</description>
*)
{endregion}
FUNCTION_BLOCK AssertInTimespan_LDT EXTENDS AssertionBase
VAR_INPUT
    IN : LDT; //! Actual value checked or observed by this Assertion.
    StartTime : LDT; //! Inclusive start of the time span; must not exceed EndTime.
    EndTime : LDT; //! Inclusive end of the time span; must not precede StartTime.
END_VAR

SUPER^();

{region 'Documentation'}
(*!
<summary>Evaluate the typed temporal relation and report higher-priority errors first.</summary>
*)
{endregion}
METHOD PROTECTED Assert
VAR
    Message : STRING(GVL_Constants.MessageLength);
    StartTimeText : STRING(GVL_Constants.AssertionValueLength);
    EndTimeText : STRING(GVL_Constants.AssertionValueLength);
    ActualText : STRING(GVL_Constants.AssertionValueLength);
END_VAR
IF NOT EvaluationActive THEN
    RETURN;
END_IF;

IF Result = E_Result.Error THEN
    RETURN;
END_IF;

IF StartTime > EndTime THEN
    StartTimeText := LDT_TO_STRING(StartTime);
    EndTimeText := LDT_TO_STRING(EndTime);
    Message := CONCAT('Assertion error: start time exceeds end time. StartTime = ',
        StartTimeText);
    Message := CONCAT(Message, ', EndTime = ');
    Message := CONCAT(Message, EndTimeText);
    Message := CONCAT(Message, '.');
    Error(Message := Message);
    RETURN;
END_IF;

IF Result = E_Result.Failed THEN
    RETURN;
END_IF;

IF (IN < StartTime) OR (IN > EndTime) THEN
    StartTimeText := LDT_TO_STRING(StartTime);
    EndTimeText := LDT_TO_STRING(EndTime);
    ActualText := LDT_TO_STRING(IN);
    Message := CONCAT('Assertion failed: value is outside allowed timespan. StartTime = ',
        StartTimeText);
    Message := CONCAT(Message, ', EndTime = ');
    Message := CONCAT(Message, EndTimeText);
    Message := CONCAT(Message, ', Actual = ');
    Message := CONCAT(Message, ActualText);
    Message := CONCAT(Message, '.');
    Fail(Message := Message);
    RETURN;
END_IF;

Pass();
END_METHOD

END_FUNCTION_BLOCK

// ---- Framework/Assertions/POU/BasicTypes/LDT/AssertLaterThan_LDT.TcPOU
{region 'Documentation'}
(*!
<summary>Check that IN is strictly later than Minimum.</summary>
*)
{endregion}
FUNCTION_BLOCK AssertLaterThan_LDT EXTENDS AssertionBase
VAR_INPUT
    IN : LDT; //! Actual value checked or observed by this Assertion.
    Minimum : LDT; //! Exclusive lower bound; the actual value or count must be greater.
END_VAR

SUPER^();

{region 'Documentation'}
(*!
<summary>Evaluate the typed temporal relation and report higher-priority errors first.</summary>
*)
{endregion}
METHOD PROTECTED Assert
VAR
    Message : STRING(GVL_Constants.MessageLength);
    MinimumText : STRING(GVL_Constants.AssertionValueLength);
    ActualText : STRING(GVL_Constants.AssertionValueLength);
END_VAR
IF NOT EvaluationActive THEN
    RETURN;
END_IF;

IF Result = E_Result.Error THEN
    RETURN;
END_IF;

IF Result = E_Result.Failed THEN
    RETURN;
END_IF;

IF IN <= Minimum THEN
    MinimumText := LDT_TO_STRING(Minimum);
    ActualText := LDT_TO_STRING(IN);
    Message := CONCAT('Assertion failed: value is not later than limit. Minimum = ',
        MinimumText);
    Message := CONCAT(Message, ', Actual = ');
    Message := CONCAT(Message, ActualText);
    Message := CONCAT(Message, '.');
    Fail(Message := Message);
    RETURN;
END_IF;

Pass();
END_METHOD

END_FUNCTION_BLOCK

// ---- Framework/Assertions/POU/BasicTypes/LDT/AssertNotEqual_LDT.TcPOU
{region 'Documentation'}
(*!
<summary>Checks inequality with the forbidden LDT value.</summary>
*)
{endregion}
FUNCTION_BLOCK AssertNotEqual_LDT EXTENDS AssertionBase
VAR_INPUT
    IN : LDT; //! Actual value checked or observed by this Assertion.
    Expected : LDT; //! Value that must differ from IN under this Assertion's comparison rules.
END_VAR

SUPER^();

{region 'Documentation'}
(*!
<summary>Evaluate the typed temporal relation and report higher-priority errors first.</summary>
*)
{endregion}
METHOD PROTECTED Assert
VAR
    Message : STRING(GVL_Constants.MessageLength);
    ExpectedText : STRING(GVL_Constants.AssertionValueLength);
    ActualText : STRING(GVL_Constants.AssertionValueLength);
END_VAR
IF NOT EvaluationActive THEN
    RETURN;
END_IF;

IF Result = E_Result.Error THEN
    RETURN;
END_IF;

IF Result = E_Result.Failed THEN
    RETURN;
END_IF;

IF IN = Expected THEN
    ExpectedText := LDT_TO_STRING(Expected);
    ActualText := LDT_TO_STRING(IN);
    Message := CONCAT('Assertion failed: values are equal but should differ. NotExpected = ',
        ExpectedText);
    Message := CONCAT(Message, ', Actual = ');
    Message := CONCAT(Message, ActualText);
    Message := CONCAT(Message, '.');
    Fail(Message := Message);
    RETURN;
END_IF;

Pass();
END_METHOD

END_FUNCTION_BLOCK

// ---- Framework/Assertions/POU/BasicTypes/LDT/AssertNotInTimespan_LDT.TcPOU
{region 'Documentation'}
(*!
<summary>Check that IN is outside the inclusive StartTime..EndTime interval.</summary>
<description>

StartTime &gt; EndTime reports Error during active evaluation; equal bounds are
valid.

</description>
*)
{endregion}
FUNCTION_BLOCK AssertNotInTimespan_LDT EXTENDS AssertionBase
VAR_INPUT
    IN : LDT; //! Actual value checked or observed by this Assertion.
    StartTime : LDT; //! Inclusive start of the time span; must not exceed EndTime.
    EndTime : LDT; //! Inclusive end of the time span; must not precede StartTime.
END_VAR

SUPER^();

{region 'Documentation'}
(*!
<summary>Evaluate the typed temporal relation and report higher-priority errors first.</summary>
*)
{endregion}
METHOD PROTECTED Assert
VAR
    Message : STRING(GVL_Constants.MessageLength);
    StartTimeText : STRING(GVL_Constants.AssertionValueLength);
    EndTimeText : STRING(GVL_Constants.AssertionValueLength);
    ActualText : STRING(GVL_Constants.AssertionValueLength);
END_VAR
IF NOT EvaluationActive THEN
    RETURN;
END_IF;

IF Result = E_Result.Error THEN
    RETURN;
END_IF;

IF StartTime > EndTime THEN
    StartTimeText := LDT_TO_STRING(StartTime);
    EndTimeText := LDT_TO_STRING(EndTime);
    Message := CONCAT('Assertion error: start time exceeds end time. StartTime = ',
        StartTimeText);
    Message := CONCAT(Message, ', EndTime = ');
    Message := CONCAT(Message, EndTimeText);
    Message := CONCAT(Message, '.');
    Error(Message := Message);
    RETURN;
END_IF;

IF Result = E_Result.Failed THEN
    RETURN;
END_IF;

IF (IN >= StartTime) AND (IN <= EndTime) THEN
    StartTimeText := LDT_TO_STRING(StartTime);
    EndTimeText := LDT_TO_STRING(EndTime);
    ActualText := LDT_TO_STRING(IN);
    Message := CONCAT('Assertion failed: value is inside forbidden timespan. StartTime = ',
        StartTimeText);
    Message := CONCAT(Message, ', EndTime = ');
    Message := CONCAT(Message, EndTimeText);
    Message := CONCAT(Message, ', Actual = ');
    Message := CONCAT(Message, ActualText);
    Message := CONCAT(Message, '.');
    Fail(Message := Message);
    RETURN;
END_IF;

Pass();
END_METHOD

END_FUNCTION_BLOCK

// ---- Framework/Assertions/POU/BasicTypes/LDT/AssertNoValueChange_LDT.TcPOU
{region 'Documentation'}
(*!
<summary>Check equality between consecutive active observations.</summary>
<description>

The first active observation establishes a baseline without deciding a result. Disabling
observation invalidates that baseline, not the held Result. Re-enabling first establishes a new
baseline; Reset clears history.

ObserveFirstCycle FALSE delays the first observation by one enabled call.

</description>
*)
{endregion}
FUNCTION_BLOCK AssertNoValueChange_LDT EXTENDS AssertionBase
VAR_INPUT
    IN : LDT; //! Actual value to observe.
END_VAR
VAR
    FINPrevious : LDT;
    FObservationPrevious : BOOL;
    FEvaluationActive : BOOL;
END_VAR

SUPER^();

{region 'Documentation'}
(*!
<summary>Observe the current value before evaluating a change against the previous observation.</summary>
*)
{endregion}
METHOD PROTECTED Assert
VAR
    PreviousValue : LDT;
    Message : STRING(GVL_Constants.MessageLength);
    PreviousText : STRING(GVL_Constants.AssertionValueLength);
    ActualText : STRING(GVL_Constants.AssertionValueLength);
END_VAR
FEvaluationActive := ObservationActive AND FObservationPrevious;
FObservationPrevious := ObservationActive;

IF NOT ObservationActive THEN
    RETURN;
END_IF;

PreviousValue := FINPrevious;
FINPrevious := IN;

IF NOT EvaluationActive THEN
    RETURN;
END_IF;

IF Result = E_Result.Error THEN
    RETURN;
END_IF;

IF Result = E_Result.Failed THEN
    RETURN;
END_IF;

IF IN <> PreviousValue THEN
    PreviousText := LDT_TO_STRING(PreviousValue);
    ActualText := LDT_TO_STRING(IN);
    Message := CONCAT('Assertion failed: value changed unexpectedly. Previous = ',
        PreviousText);
    Message := CONCAT(Message, ', Actual = ');
    Message := CONCAT(Message, ActualText);
    Message := CONCAT(Message, '.');
    Fail(Message := Message);
    RETURN;
END_IF;

Pass();
END_METHOD

{region 'Documentation'}
(*!
<summary>Current/last call has an active observation and a preceding observation
baseline.</summary>
*)
{endregion}
{attribute 'monitoring' := 'call'}
PROPERTY PUBLIC EvaluationActive : BOOL //! Current/last call has an active observation and a preceding observation baseline.
GET // PUBLIC
EvaluationActive := FEvaluationActive;
END_GET
END_PROPERTY

{region 'Documentation'}
(*!
<summary>Clear observation history and the current evaluation gate.</summary>
*)
{endregion}
METHOD PROTECTED ResetAssertion
FINPrevious := LDT#1970-01-01-00:00:00;
FObservationPrevious := FALSE;
FEvaluationActive := FALSE;
END_METHOD

END_FUNCTION_BLOCK

// ---- Framework/Assertions/POU/BasicTypes/LInt/AssertNoValueChange_LInt.TcPOU
{region 'Documentation'}
(*!
<summary>Check equality between consecutive active observations.</summary>
<description>

The first active observation establishes a baseline without deciding a result. Disabling
observation invalidates that baseline, not the held Result. Re-enabling first establishes a new
baseline; Reset clears history.

ObserveFirstCycle FALSE delays the first observation by one enabled call.

</description>
*)
{endregion}
FUNCTION_BLOCK AssertNoValueChange_LInt EXTENDS AssertionBase
VAR_INPUT
    IN : LINT; //! Actual value to observe.
END_VAR
VAR
    FINPrevious : LINT;
    FObservationPrevious : BOOL;
    FEvaluationActive : BOOL;
END_VAR

SUPER^();

{region 'Documentation'}
(*!
<summary>Observe the current value before evaluating a change against the previous observation.</summary>
*)
{endregion}
METHOD PROTECTED Assert
VAR
    PreviousValue : LINT;
    Message : STRING(GVL_Constants.MessageLength);
    PreviousText : STRING(GVL_Constants.AssertionValueLength);
    ActualText : STRING(GVL_Constants.AssertionValueLength);
END_VAR
FEvaluationActive := ObservationActive AND FObservationPrevious;
FObservationPrevious := ObservationActive;

IF NOT ObservationActive THEN
    RETURN;
END_IF;

PreviousValue := FINPrevious;
FINPrevious := IN;

IF NOT EvaluationActive THEN
    RETURN;
END_IF;

IF Result = E_Result.Error THEN
    RETURN;
END_IF;

IF Result = E_Result.Failed THEN
    RETURN;
END_IF;

IF IN <> PreviousValue THEN
    PreviousText := LINT_TO_STRING(PreviousValue);
    ActualText := LINT_TO_STRING(IN);
    Message := CONCAT('Assertion failed: value changed unexpectedly. Previous = ',
        PreviousText);
    Message := CONCAT(Message, ', Actual = ');
    Message := CONCAT(Message, ActualText);
    Message := CONCAT(Message, '.');
    Fail(Message := Message);
    RETURN;
END_IF;

Pass();
END_METHOD

{region 'Documentation'}
(*!
<summary>Current/last call has an active observation and a preceding observation
baseline.</summary>
*)
{endregion}
{attribute 'monitoring' := 'call'}
PROPERTY PUBLIC EvaluationActive : BOOL //! Current/last call has an active observation and a preceding observation baseline.
GET // PUBLIC
EvaluationActive := FEvaluationActive;
END_GET
END_PROPERTY

{region 'Documentation'}
(*!
<summary>Clear observation history and the current evaluation gate.</summary>
*)
{endregion}
METHOD PROTECTED ResetAssertion
FINPrevious := 0;
FObservationPrevious := FALSE;
FEvaluationActive := FALSE;
END_METHOD

END_FUNCTION_BLOCK

// ---- Framework/Assertions/POU/BasicTypes/LInt/AssertSequence_LInt.TcPOU
{region 'Documentation'}
(*!
<summary>Checks the observed value sequence; Evaluate also checks the current value and
completeness.</summary>
<description>

Uses the whole Expected array from its declared lower bound. Keep its binding, bounds and
values stable until Reset; supply it on reset and disabled FB calls as well.

Observation accepts the current expected value and then permits advancing by one element
on a later change. Repeated equal values do not advance. An unexpected value or an out-of-range
sequence index reports Failed.

Evaluate checks the current value and requires the final expected element to have been
reached; only then can the result become Passed. Disabling observation retains progression.
Reset restarts it.

</description>
*)
{endregion}
FUNCTION_BLOCK AssertSequence_LInt EXTENDS AssertionWithEvaluationBase
VAR_INPUT
    IN : LINT; //! Actual value to observe.
END_VAR
VAR_IN_OUT CONSTANT
    Expected : ARRAY[*] OF LINT; //! Complete expected sequence; read without modifying the supplied array.
END_VAR
VAR
    FExpectedIndex : DINT;
    FSequenceIndexInitialized : BOOL;
    FAllowAdvance : BOOL;
END_VAR

SUPER^();

{region 'Documentation'}
(*!
<summary>Advances at most one entry and checks the current value before explicit completeness evaluation.</summary>
*)
{endregion}
METHOD PROTECTED Assert
VAR
    LowerIndex : DINT;
    UpperIndex : DINT;
    ExpectedValue : LINT;
    MatchesExpected : BOOL;
    AllowAdvance : BOOL;
    Message : STRING(GVL_Constants.MessageLength);
    ExpectedText : STRING(GVL_Constants.AssertionValueLength);
    ActualText : STRING(GVL_Constants.AssertionValueLength);
END_VAR
LowerIndex := LOWER_BOUND(Expected, 1);
UpperIndex := UPPER_BOUND(Expected, 1);

IF NOT FSequenceIndexInitialized THEN
    FExpectedIndex := LowerIndex;
    FSequenceIndexInitialized := TRUE;
END_IF;

IF NOT (ObservationActive OR EvaluationActive) THEN
    RETURN;
END_IF;

IF Result = E_Result.Error THEN
    RETURN;
END_IF;

IF Result = E_Result.Failed THEN
    RETURN;
END_IF;

IF (FExpectedIndex < LowerIndex) OR (FExpectedIndex > UpperIndex) THEN
    Message := CONCAT('Assertion failed: sequence index out of range. ExpectedIndex = ',
        DINT_TO_STRING(FExpectedIndex));
    Message := CONCAT(Message, ', LowerIndex = ');
    Message := CONCAT(Message, DINT_TO_STRING(LowerIndex));
    Message := CONCAT(Message, ', UpperIndex = ');
    Message := CONCAT(Message, DINT_TO_STRING(UpperIndex));
    Message := CONCAT(Message, '.');
    Fail(Message := Message);
    RETURN;
END_IF;

AllowAdvance := FAllowAdvance;
IF ObservationActive THEN
    FAllowAdvance := TRUE;
END_IF;

ExpectedValue := Expected[FExpectedIndex];
MatchesExpected := IN = ExpectedValue;

IF AllowAdvance AND NOT MatchesExpected THEN
    IF FExpectedIndex = UpperIndex THEN
        Message := CONCAT('Assertion failed: sequence continued beyond its last entry. LastIndex = ',
            DINT_TO_STRING(UpperIndex));
        Message := CONCAT(Message, '.');
        Fail(Message := Message);
        RETURN;
    END_IF;

    FExpectedIndex := FExpectedIndex + 1;
    ExpectedValue := Expected[FExpectedIndex];
    MatchesExpected := IN = ExpectedValue;
END_IF;

IF NOT MatchesExpected THEN
    ExpectedText := LINT_TO_STRING(ExpectedValue);
    ActualText := LINT_TO_STRING(IN);
    Message := CONCAT('Assertion failed: sequence value does not match. ExpectedIndex = ',
        DINT_TO_STRING(FExpectedIndex));
    Message := CONCAT(Message, ', Expected = ');
    Message := CONCAT(Message, ExpectedText);
    Message := CONCAT(Message, ', Actual = ');
    Message := CONCAT(Message, ActualText);
    Message := CONCAT(Message, '.');
    Fail(Message := Message);
    RETURN;
END_IF;

IF NOT EvaluationActive THEN
    RETURN;
END_IF;

IF FExpectedIndex <> UpperIndex THEN
    Message := CONCAT('Assertion failed: sequence is incomplete. ExpectedIndex = ',
        DINT_TO_STRING(FExpectedIndex));
    Message := CONCAT(Message, ', LastIndex = ');
    Message := CONCAT(Message, DINT_TO_STRING(UpperIndex));
    Message := CONCAT(Message, '.');
    Fail(Message := Message);
    RETURN;
END_IF;

Pass();
END_METHOD

{region 'Documentation'}
(*!
<summary>Restart progression at the bound Expected array's lower index.</summary>
<description>

Runs only during the reset FB call with Expected supplied, not directly from Reset or
Initialize. Clears permission to advance from a previous observation.

</description>
*)
{endregion}
METHOD PROTECTED ResetAssertion
FExpectedIndex := LOWER_BOUND(Expected, 1);
FSequenceIndexInitialized := TRUE;
FAllowAdvance := FALSE;
END_METHOD

END_FUNCTION_BLOCK

// ---- Framework/Assertions/POU/BasicTypes/LTime/AssertEarlierThan_LTime.TcPOU
{region 'Documentation'}
(*!
<summary>Check that IN is strictly earlier than Maximum.</summary>
*)
{endregion}
FUNCTION_BLOCK AssertEarlierThan_LTime EXTENDS AssertionBase
VAR_INPUT
    IN : LTIME; //! Actual value checked or observed by this Assertion.
    Maximum : LTIME; //! Exclusive upper bound; the actual value or count must be smaller.
END_VAR

SUPER^();

{region 'Documentation'}
(*!
<summary>Evaluate the typed duration relation and report higher-priority errors first.</summary>
*)
{endregion}
METHOD PROTECTED Assert
VAR
    Message : STRING(GVL_Constants.MessageLength);
    MaximumText : STRING(GVL_Constants.AssertionValueLength);
    ActualText : STRING(GVL_Constants.AssertionValueLength);
END_VAR
IF NOT EvaluationActive THEN
    RETURN;
END_IF;

IF Result = E_Result.Error THEN
    RETURN;
END_IF;

IF Result = E_Result.Failed THEN
    RETURN;
END_IF;

IF IN >= Maximum THEN
    MaximumText := LTIME_TO_STRING(Maximum);
    ActualText := LTIME_TO_STRING(IN);
    Message := CONCAT('Assertion failed: value is not earlier than limit. Maximum = ',
        MaximumText);
    Message := CONCAT(Message, ', Actual = ');
    Message := CONCAT(Message, ActualText);
    Message := CONCAT(Message, '.');
    Fail(Message := Message);
    RETURN;
END_IF;

Pass();
END_METHOD

END_FUNCTION_BLOCK

// ---- Framework/Assertions/POU/BasicTypes/LTime/AssertInTimespan_LTime.TcPOU
{region 'Documentation'}
(*!
<summary>Check that IN is inside the inclusive StartTime..EndTime interval.</summary>
<description>

StartTime &gt; EndTime reports Error during active evaluation; equal bounds are
valid.

</description>
*)
{endregion}
FUNCTION_BLOCK AssertInTimespan_LTime EXTENDS AssertionBase
VAR_INPUT
    IN : LTIME; //! Actual value checked or observed by this Assertion.
    StartTime : LTIME; //! Inclusive start of the time span; must not exceed EndTime.
    EndTime : LTIME; //! Inclusive end of the time span; must not precede StartTime.
END_VAR

SUPER^();

{region 'Documentation'}
(*!
<summary>Evaluate the typed duration relation and report higher-priority errors first.</summary>
*)
{endregion}
METHOD PROTECTED Assert
VAR
    Message : STRING(GVL_Constants.MessageLength);
    StartTimeText : STRING(GVL_Constants.AssertionValueLength);
    EndTimeText : STRING(GVL_Constants.AssertionValueLength);
    ActualText : STRING(GVL_Constants.AssertionValueLength);
END_VAR
IF NOT EvaluationActive THEN
    RETURN;
END_IF;

IF Result = E_Result.Error THEN
    RETURN;
END_IF;

IF StartTime > EndTime THEN
    StartTimeText := LTIME_TO_STRING(StartTime);
    EndTimeText := LTIME_TO_STRING(EndTime);
    Message := CONCAT('Assertion error: start time exceeds end time. StartTime = ',
        StartTimeText);
    Message := CONCAT(Message, ', EndTime = ');
    Message := CONCAT(Message, EndTimeText);
    Message := CONCAT(Message, '.');
    Error(Message := Message);
    RETURN;
END_IF;

IF Result = E_Result.Failed THEN
    RETURN;
END_IF;

IF (IN < StartTime) OR (IN > EndTime) THEN
    StartTimeText := LTIME_TO_STRING(StartTime);
    EndTimeText := LTIME_TO_STRING(EndTime);
    ActualText := LTIME_TO_STRING(IN);
    Message := CONCAT('Assertion failed: value is outside allowed timespan. StartTime = ',
        StartTimeText);
    Message := CONCAT(Message, ', EndTime = ');
    Message := CONCAT(Message, EndTimeText);
    Message := CONCAT(Message, ', Actual = ');
    Message := CONCAT(Message, ActualText);
    Message := CONCAT(Message, '.');
    Fail(Message := Message);
    RETURN;
END_IF;

Pass();
END_METHOD

END_FUNCTION_BLOCK

// ---- Framework/Assertions/POU/BasicTypes/LTime/AssertLaterThan_LTime.TcPOU
{region 'Documentation'}
(*!
<summary>Check that IN is strictly later than Minimum.</summary>
*)
{endregion}
FUNCTION_BLOCK AssertLaterThan_LTime EXTENDS AssertionBase
VAR_INPUT
    IN : LTIME; //! Actual value checked or observed by this Assertion.
    Minimum : LTIME; //! Exclusive lower bound; the actual value or count must be greater.
END_VAR

SUPER^();

{region 'Documentation'}
(*!
<summary>Evaluate the typed duration relation and report higher-priority errors first.</summary>
*)
{endregion}
METHOD PROTECTED Assert
VAR
    Message : STRING(GVL_Constants.MessageLength);
    MinimumText : STRING(GVL_Constants.AssertionValueLength);
    ActualText : STRING(GVL_Constants.AssertionValueLength);
END_VAR
IF NOT EvaluationActive THEN
    RETURN;
END_IF;

IF Result = E_Result.Error THEN
    RETURN;
END_IF;

IF Result = E_Result.Failed THEN
    RETURN;
END_IF;

IF IN <= Minimum THEN
    MinimumText := LTIME_TO_STRING(Minimum);
    ActualText := LTIME_TO_STRING(IN);
    Message := CONCAT('Assertion failed: value is not later than limit. Minimum = ',
        MinimumText);
    Message := CONCAT(Message, ', Actual = ');
    Message := CONCAT(Message, ActualText);
    Message := CONCAT(Message, '.');
    Fail(Message := Message);
    RETURN;
END_IF;

Pass();
END_METHOD

END_FUNCTION_BLOCK

// ---- Framework/Assertions/POU/BasicTypes/LTime/AssertNotEqual_LTime.TcPOU
{region 'Documentation'}
(*!
<summary>Checks inequality with the forbidden LTIME value.</summary>
*)
{endregion}
FUNCTION_BLOCK AssertNotEqual_LTime EXTENDS AssertionBase
VAR_INPUT
    IN : LTIME; //! Actual value checked or observed by this Assertion.
    Expected : LTIME; //! Value that must differ from IN under this Assertion's comparison rules.
END_VAR

SUPER^();

{region 'Documentation'}
(*!
<summary>Evaluate the typed duration relation and report higher-priority errors first.</summary>
*)
{endregion}
METHOD PROTECTED Assert
VAR
    Message : STRING(GVL_Constants.MessageLength);
    ExpectedText : STRING(GVL_Constants.AssertionValueLength);
    ActualText : STRING(GVL_Constants.AssertionValueLength);
END_VAR
IF NOT EvaluationActive THEN
    RETURN;
END_IF;

IF Result = E_Result.Error THEN
    RETURN;
END_IF;

IF Result = E_Result.Failed THEN
    RETURN;
END_IF;

IF IN = Expected THEN
    ExpectedText := LTIME_TO_STRING(Expected);
    ActualText := LTIME_TO_STRING(IN);
    Message := CONCAT('Assertion failed: values are equal but should differ. NotExpected = ',
        ExpectedText);
    Message := CONCAT(Message, ', Actual = ');
    Message := CONCAT(Message, ActualText);
    Message := CONCAT(Message, '.');
    Fail(Message := Message);
    RETURN;
END_IF;

Pass();
END_METHOD

END_FUNCTION_BLOCK

// ---- Framework/Assertions/POU/BasicTypes/LTime/AssertNotInTimespan_LTime.TcPOU
{region 'Documentation'}
(*!
<summary>Check that IN is outside the inclusive StartTime..EndTime interval.</summary>
<description>

StartTime &gt; EndTime reports Error during active evaluation; equal bounds are
valid.

</description>
*)
{endregion}
FUNCTION_BLOCK AssertNotInTimespan_LTime EXTENDS AssertionBase
VAR_INPUT
    IN : LTIME; //! Actual value checked or observed by this Assertion.
    StartTime : LTIME; //! Inclusive start of the time span; must not exceed EndTime.
    EndTime : LTIME; //! Inclusive end of the time span; must not precede StartTime.
END_VAR

SUPER^();

{region 'Documentation'}
(*!
<summary>Evaluate the typed duration relation and report higher-priority errors first.</summary>
*)
{endregion}
METHOD PROTECTED Assert
VAR
    Message : STRING(GVL_Constants.MessageLength);
    StartTimeText : STRING(GVL_Constants.AssertionValueLength);
    EndTimeText : STRING(GVL_Constants.AssertionValueLength);
    ActualText : STRING(GVL_Constants.AssertionValueLength);
END_VAR
IF NOT EvaluationActive THEN
    RETURN;
END_IF;

IF Result = E_Result.Error THEN
    RETURN;
END_IF;

IF StartTime > EndTime THEN
    StartTimeText := LTIME_TO_STRING(StartTime);
    EndTimeText := LTIME_TO_STRING(EndTime);
    Message := CONCAT('Assertion error: start time exceeds end time. StartTime = ',
        StartTimeText);
    Message := CONCAT(Message, ', EndTime = ');
    Message := CONCAT(Message, EndTimeText);
    Message := CONCAT(Message, '.');
    Error(Message := Message);
    RETURN;
END_IF;

IF Result = E_Result.Failed THEN
    RETURN;
END_IF;

IF (IN >= StartTime) AND (IN <= EndTime) THEN
    StartTimeText := LTIME_TO_STRING(StartTime);
    EndTimeText := LTIME_TO_STRING(EndTime);
    ActualText := LTIME_TO_STRING(IN);
    Message := CONCAT('Assertion failed: value is inside forbidden timespan. StartTime = ',
        StartTimeText);
    Message := CONCAT(Message, ', EndTime = ');
    Message := CONCAT(Message, EndTimeText);
    Message := CONCAT(Message, ', Actual = ');
    Message := CONCAT(Message, ActualText);
    Message := CONCAT(Message, '.');
    Fail(Message := Message);
    RETURN;
END_IF;

Pass();
END_METHOD

END_FUNCTION_BLOCK

// ---- Framework/Assertions/POU/BasicTypes/LTime/AssertNoValueChange_LTime.TcPOU
{region 'Documentation'}
(*!
<summary>Check equality between consecutive active observations.</summary>
<description>

The first active observation establishes a baseline without deciding a result. Disabling
observation invalidates that baseline, not the held Result. Re-enabling first establishes a new
baseline; Reset clears history.

ObserveFirstCycle FALSE delays the first observation by one enabled call.

</description>
*)
{endregion}
FUNCTION_BLOCK AssertNoValueChange_LTime EXTENDS AssertionBase
VAR_INPUT
    IN : LTIME; //! Actual value to observe.
END_VAR
VAR
    FINPrevious : LTIME;
    FObservationPrevious : BOOL;
    FEvaluationActive : BOOL;
END_VAR

SUPER^();

{region 'Documentation'}
(*!
<summary>Observe the current value before evaluating a change against the previous observation.</summary>
*)
{endregion}
METHOD PROTECTED Assert
VAR
    PreviousValue : LTIME;
    Message : STRING(GVL_Constants.MessageLength);
    PreviousText : STRING(GVL_Constants.AssertionValueLength);
    ActualText : STRING(GVL_Constants.AssertionValueLength);
END_VAR
FEvaluationActive := ObservationActive AND FObservationPrevious;
FObservationPrevious := ObservationActive;

IF NOT ObservationActive THEN
    RETURN;
END_IF;

PreviousValue := FINPrevious;
FINPrevious := IN;

IF NOT EvaluationActive THEN
    RETURN;
END_IF;

IF Result = E_Result.Error THEN
    RETURN;
END_IF;

IF Result = E_Result.Failed THEN
    RETURN;
END_IF;

IF IN <> PreviousValue THEN
    PreviousText := LTIME_TO_STRING(PreviousValue);
    ActualText := LTIME_TO_STRING(IN);
    Message := CONCAT('Assertion failed: value changed unexpectedly. Previous = ',
        PreviousText);
    Message := CONCAT(Message, ', Actual = ');
    Message := CONCAT(Message, ActualText);
    Message := CONCAT(Message, '.');
    Fail(Message := Message);
    RETURN;
END_IF;

Pass();
END_METHOD

{region 'Documentation'}
(*!
<summary>Current/last call has an active observation and a preceding observation
baseline.</summary>
*)
{endregion}
{attribute 'monitoring' := 'call'}
PROPERTY PUBLIC EvaluationActive : BOOL //! Current/last call has an active observation and a preceding observation baseline.
GET // PUBLIC
EvaluationActive := FEvaluationActive;
END_GET
END_PROPERTY

{region 'Documentation'}
(*!
<summary>Clear observation history and the current evaluation gate.</summary>
*)
{endregion}
METHOD PROTECTED ResetAssertion
FINPrevious := LTIME#0ns;
FObservationPrevious := FALSE;
FEvaluationActive := FALSE;
END_METHOD

END_FUNCTION_BLOCK

// ---- Framework/Assertions/POU/BasicTypes/LTOD/AssertEarlierThan_LTOD.TcPOU
{region 'Documentation'}
(*!
<summary>Check that IN is strictly earlier than Maximum.</summary>
<description>

A value at or beyond 24 hours reports Error before comparison or baseline capture.

</description>
*)
{endregion}
FUNCTION_BLOCK AssertEarlierThan_LTOD EXTENDS AssertionBase
VAR_INPUT
    IN : LTOD; //! Actual value checked or observed by this Assertion.
    Maximum : LTOD; //! Exclusive upper bound; the actual value or count must be smaller.
END_VAR

SUPER^();

{region 'Documentation'}
(*!
<summary>Evaluate the typed temporal relation and report higher-priority errors first.</summary>
*)
{endregion}
METHOD PROTECTED Assert
VAR
    Message : STRING(GVL_Constants.MessageLength);
    MaximumText : STRING(GVL_Constants.AssertionValueLength);
    ActualText : STRING(GVL_Constants.AssertionValueLength);
END_VAR
IF NOT EvaluationActive THEN
    RETURN;
END_IF;

IF Result = E_Result.Error THEN
    RETURN;
END_IF;

IF NOT IsTimeOfDayValid_LTOD(Value := IN) THEN
    Error(Message := 'Assertion error: IN is outside the valid LTOD range (less than 24 hours).');
    RETURN;
END_IF;

IF NOT IsTimeOfDayValid_LTOD(Value := Maximum) THEN
    Error(Message := 'Assertion error: Maximum is outside the valid LTOD range (less than 24 hours).');
    RETURN;
END_IF;

IF Result = E_Result.Failed THEN
    RETURN;
END_IF;

IF IN >= Maximum THEN
    MaximumText := LTOD_TO_STRING(Maximum);
    ActualText := LTOD_TO_STRING(IN);
    Message := CONCAT('Assertion failed: value is not earlier than limit. Maximum = ',
        MaximumText);
    Message := CONCAT(Message, ', Actual = ');
    Message := CONCAT(Message, ActualText);
    Message := CONCAT(Message, '.');
    Fail(Message := Message);
    RETURN;
END_IF;

Pass();
END_METHOD

END_FUNCTION_BLOCK

// ---- Framework/Assertions/POU/BasicTypes/LTOD/AssertLaterThan_LTOD.TcPOU
{region 'Documentation'}
(*!
<summary>Check that IN is strictly later than Minimum.</summary>
<description>

A value at or beyond 24 hours reports Error before comparison or baseline capture.

</description>
*)
{endregion}
FUNCTION_BLOCK AssertLaterThan_LTOD EXTENDS AssertionBase
VAR_INPUT
    IN : LTOD; //! Actual value checked or observed by this Assertion.
    Minimum : LTOD; //! Exclusive lower bound; the actual value or count must be greater.
END_VAR

SUPER^();

{region 'Documentation'}
(*!
<summary>Evaluate the typed temporal relation and report higher-priority errors first.</summary>
*)
{endregion}
METHOD PROTECTED Assert
VAR
    Message : STRING(GVL_Constants.MessageLength);
    MinimumText : STRING(GVL_Constants.AssertionValueLength);
    ActualText : STRING(GVL_Constants.AssertionValueLength);
END_VAR
IF NOT EvaluationActive THEN
    RETURN;
END_IF;

IF Result = E_Result.Error THEN
    RETURN;
END_IF;

IF NOT IsTimeOfDayValid_LTOD(Value := IN) THEN
    Error(Message := 'Assertion error: IN is outside the valid LTOD range (less than 24 hours).');
    RETURN;
END_IF;

IF NOT IsTimeOfDayValid_LTOD(Value := Minimum) THEN
    Error(Message := 'Assertion error: Minimum is outside the valid LTOD range (less than 24 hours).');
    RETURN;
END_IF;

IF Result = E_Result.Failed THEN
    RETURN;
END_IF;

IF IN <= Minimum THEN
    MinimumText := LTOD_TO_STRING(Minimum);
    ActualText := LTOD_TO_STRING(IN);
    Message := CONCAT('Assertion failed: value is not later than limit. Minimum = ',
        MinimumText);
    Message := CONCAT(Message, ', Actual = ');
    Message := CONCAT(Message, ActualText);
    Message := CONCAT(Message, '.');
    Fail(Message := Message);
    RETURN;
END_IF;

Pass();
END_METHOD

END_FUNCTION_BLOCK

// ---- Framework/Assertions/POU/BasicTypes/LTOD/AssertNotEqual_LTOD.TcPOU
{region 'Documentation'}
(*!
<summary>Checks inequality with the forbidden LTOD value.</summary>
<description>

A value at or beyond 24 hours reports Error before comparison or baseline capture.

</description>
*)
{endregion}
FUNCTION_BLOCK AssertNotEqual_LTOD EXTENDS AssertionBase
VAR_INPUT
    IN : LTOD; //! Actual value checked or observed by this Assertion.
    Expected : LTOD; //! Value that must differ from IN under this Assertion's comparison rules.
END_VAR

SUPER^();

{region 'Documentation'}
(*!
<summary>Evaluate the typed temporal relation and report higher-priority errors first.</summary>
*)
{endregion}
METHOD PROTECTED Assert
VAR
    Message : STRING(GVL_Constants.MessageLength);
    ExpectedText : STRING(GVL_Constants.AssertionValueLength);
    ActualText : STRING(GVL_Constants.AssertionValueLength);
END_VAR
IF NOT EvaluationActive THEN
    RETURN;
END_IF;

IF Result = E_Result.Error THEN
    RETURN;
END_IF;

IF NOT IsTimeOfDayValid_LTOD(Value := IN) THEN
    Error(Message := 'Assertion error: IN is outside the valid LTOD range (less than 24 hours).');
    RETURN;
END_IF;

IF NOT IsTimeOfDayValid_LTOD(Value := Expected) THEN
    Error(Message := 'Assertion error: Expected is outside the valid LTOD range (less than 24 hours).');
    RETURN;
END_IF;

IF Result = E_Result.Failed THEN
    RETURN;
END_IF;

IF IN = Expected THEN
    ExpectedText := LTOD_TO_STRING(Expected);
    ActualText := LTOD_TO_STRING(IN);
    Message := CONCAT('Assertion failed: values are equal but should differ. NotExpected = ',
        ExpectedText);
    Message := CONCAT(Message, ', Actual = ');
    Message := CONCAT(Message, ActualText);
    Message := CONCAT(Message, '.');
    Fail(Message := Message);
    RETURN;
END_IF;

Pass();
END_METHOD

END_FUNCTION_BLOCK

// ---- Framework/Assertions/POU/BasicTypes/LTOD/AssertNoValueChange_LTOD.TcPOU
{region 'Documentation'}
(*!
<summary>Check equality between consecutive active observations.</summary>
<description>

The first active observation establishes a baseline without deciding a result. Disabling
observation invalidates that baseline, not the held Result. Re-enabling first establishes a new
baseline; Reset clears history.

ObserveFirstCycle FALSE delays the first observation by one enabled call.

An observed value at or beyond 24 hours reports Error, including baseline capture.

</description>
*)
{endregion}
FUNCTION_BLOCK AssertNoValueChange_LTOD EXTENDS AssertionBase
VAR_INPUT
    IN : LTOD; //! Actual value to observe.
END_VAR
VAR
    FINPrevious : LTOD;
    FObservationPrevious : BOOL;
    FEvaluationActive : BOOL;
END_VAR

SUPER^();

{region 'Documentation'}
(*!
<summary>Observe the current value before evaluating a change against the previous observation.</summary>
*)
{endregion}
METHOD PROTECTED Assert
VAR
    PreviousValue : LTOD;
    Message : STRING(GVL_Constants.MessageLength);
    PreviousText : STRING(GVL_Constants.AssertionValueLength);
    ActualText : STRING(GVL_Constants.AssertionValueLength);
END_VAR
FEvaluationActive := ObservationActive AND FObservationPrevious;
FObservationPrevious := ObservationActive;

IF NOT ObservationActive THEN
    RETURN;
END_IF;

IF Result = E_Result.Error THEN
    RETURN;
END_IF;

IF NOT IsTimeOfDayValid_LTOD(Value := IN) THEN
    Error(Message := 'Assertion error: IN is outside the valid LTOD range (less than 24 hours).');
    RETURN;
END_IF;

PreviousValue := FINPrevious;
FINPrevious := IN;

IF NOT EvaluationActive THEN
    RETURN;
END_IF;

IF Result = E_Result.Failed THEN
    RETURN;
END_IF;

IF IN <> PreviousValue THEN
    PreviousText := LTOD_TO_STRING(PreviousValue);
    ActualText := LTOD_TO_STRING(IN);
    Message := CONCAT('Assertion failed: value changed unexpectedly. Previous = ',
        PreviousText);
    Message := CONCAT(Message, ', Actual = ');
    Message := CONCAT(Message, ActualText);
    Message := CONCAT(Message, '.');
    Fail(Message := Message);
    RETURN;
END_IF;

Pass();
END_METHOD

{region 'Documentation'}
(*!
<summary>Current/last call has an active observation and a preceding observation
baseline.</summary>
*)
{endregion}
{attribute 'monitoring' := 'call'}
PROPERTY PUBLIC EvaluationActive : BOOL //! Current/last call has an active observation and a preceding observation baseline.
GET // PUBLIC
EvaluationActive := FEvaluationActive;
END_GET
END_PROPERTY

{region 'Documentation'}
(*!
<summary>Clear observation history and the current evaluation gate.</summary>
*)
{endregion}
METHOD PROTECTED ResetAssertion
FINPrevious := LTOD#00:00:00;
FObservationPrevious := FALSE;
FEvaluationActive := FALSE;
END_METHOD

END_FUNCTION_BLOCK

// ---- Framework/Assertions/POU/BasicTypes/LWord/AssertContainsFalse_LWord.TcPOU
{region 'Documentation'}
(*!
<summary>Checks that at least one selected bit is FALSE.</summary>
*)
{endregion}
FUNCTION_BLOCK AssertContainsFalse_LWord EXTENDS AssertionBase
VAR_INPUT
    IN : LWORD; //! Actual bitfield.
    Mask : LWORD := 16#FFFFFFFFFFFFFFFF; //! Selects evaluated bits; defaults to all bits. An empty mask produces Error during evaluation.
END_VAR

SUPER^();

{region 'Documentation'}
(*!
<summary>Rejects an empty mask before checking for a matching selected bit.</summary>
*)
{endregion}
METHOD PROTECTED Assert
VAR
    Message : STRING(GVL_Constants.MessageLength);
    MaskText : STRING(GVL_Constants.AssertionValueLength);
    ActualText : STRING(GVL_Constants.AssertionValueLength);
END_VAR
VAR CONSTANT
    NoMask : LWORD := 16#00;
    HexDigitCount : USINT := 16;
END_VAR
IF NOT EvaluationActive THEN
    RETURN;
END_IF;

IF Result = E_Result.Error THEN
    RETURN;
END_IF;

IF Mask = NoMask THEN
    MaskText := CreateAssertionTextValue_Hex(Value := Mask,
        DigitCount := HexDigitCount);
    Message := CONCAT('Assertion error: mask must not be empty. Mask = ',
        MaskText);
    Message := CONCAT(Message, '.');
    Error(Message := Message);
    RETURN;
END_IF;

IF Result = E_Result.Failed THEN
    RETURN;
END_IF;

IF (IN AND Mask) = Mask THEN
    MaskText := CreateAssertionTextValue_Hex(Value := Mask,
        DigitCount := HexDigitCount);
    ActualText := CreateAssertionTextValue_Hex(Value := IN,
        DigitCount := HexDigitCount);
    Message := CONCAT('Assertion failed: no selected bit is FALSE. Mask = ',
        MaskText);
    Message := CONCAT(Message, ', Actual = ');
    Message := CONCAT(Message, ActualText);
    Message := CONCAT(Message, '.');
    Fail(Message := Message);
    RETURN;
END_IF;

Pass();
END_METHOD

END_FUNCTION_BLOCK

// ---- Framework/Assertions/POU/BasicTypes/LWord/AssertContainsTrue_LWord.TcPOU
{region 'Documentation'}
(*!
<summary>Checks that at least one selected bit is TRUE.</summary>
*)
{endregion}
FUNCTION_BLOCK AssertContainsTrue_LWord EXTENDS AssertionBase
VAR_INPUT
    IN : LWORD; //! Actual bitfield.
    Mask : LWORD := 16#FFFFFFFFFFFFFFFF; //! Selects evaluated bits; defaults to all bits. An empty mask produces Error during evaluation.
END_VAR

SUPER^();

{region 'Documentation'}
(*!
<summary>Rejects an empty mask before checking for a matching selected bit.</summary>
*)
{endregion}
METHOD PROTECTED Assert
VAR
    Message : STRING(GVL_Constants.MessageLength);
    MaskText : STRING(GVL_Constants.AssertionValueLength);
    ActualText : STRING(GVL_Constants.AssertionValueLength);
END_VAR
VAR CONSTANT
    NoMask : LWORD := 16#00;
    HexDigitCount : USINT := 16;
END_VAR
IF NOT EvaluationActive THEN
    RETURN;
END_IF;

IF Result = E_Result.Error THEN
    RETURN;
END_IF;

IF Mask = NoMask THEN
    MaskText := CreateAssertionTextValue_Hex(Value := Mask,
        DigitCount := HexDigitCount);
    Message := CONCAT('Assertion error: mask must not be empty. Mask = ',
        MaskText);
    Message := CONCAT(Message, '.');
    Error(Message := Message);
    RETURN;
END_IF;

IF Result = E_Result.Failed THEN
    RETURN;
END_IF;

IF (IN AND Mask) = NoMask THEN
    MaskText := CreateAssertionTextValue_Hex(Value := Mask,
        DigitCount := HexDigitCount);
    ActualText := CreateAssertionTextValue_Hex(Value := IN,
        DigitCount := HexDigitCount);
    Message := CONCAT('Assertion failed: no selected bit is TRUE. Mask = ',
        MaskText);
    Message := CONCAT(Message, ', Actual = ');
    Message := CONCAT(Message, ActualText);
    Message := CONCAT(Message, '.');
    Fail(Message := Message);
    RETURN;
END_IF;

Pass();
END_METHOD

END_FUNCTION_BLOCK

// ---- Framework/Assertions/POU/BasicTypes/LWord/AssertEqualBit_LWord.TcPOU
{region 'Documentation'}
(*!
<summary>Checks that the selected LWORD bit equals the expected Boolean value.</summary>
*)
{endregion}
FUNCTION_BLOCK AssertEqualBit_LWord EXTENDS AssertionBase
VAR_INPUT
    IN : LWORD; //! Actual bitfield.
    BitIndex : USINT; //! Zero-based bit index (0..63); an invalid index produces Error during evaluation.
    Expected : BOOL; //! Expected selected bit value.
END_VAR

SUPER^();

{region 'Documentation'}
(*!
<summary>Validates the index before evaluating the selected bit.</summary>
*)
{endregion}
METHOD PROTECTED Assert
VAR
    Mask : LWORD;
    ActualBit : BOOL;
    Message : STRING(GVL_Constants.MessageLength);
    ActualText : STRING(GVL_Constants.AssertionValueLength);
END_VAR
VAR CONSTANT
    MaxBitIndex : USINT := 63;
    SingleBitMask : LWORD := 16#01;
    NoBitMask : LWORD := 16#00;
    HexDigitCount : USINT := 16;
END_VAR
IF NOT EvaluationActive THEN
    RETURN;
END_IF;

IF Result = E_Result.Error THEN
    RETURN;
END_IF;

IF BitIndex > MaxBitIndex THEN
    Message := CONCAT('Assertion error: bit index is outside valid range. BitIndex = ',
        USINT_TO_STRING(BitIndex));
    Message := CONCAT(Message, ', MaxBitIndex = ');
    Message := CONCAT(Message, USINT_TO_STRING(MaxBitIndex));
    Message := CONCAT(Message, '.');
    Error(Message := Message);
    RETURN;
END_IF;

IF Result = E_Result.Failed THEN
    RETURN;
END_IF;

Mask := SHL(SingleBitMask, BitIndex);
ActualBit := (IN AND Mask) <> NoBitMask;

IF ActualBit <> Expected THEN
    ActualText := CreateAssertionTextValue_Hex(Value := IN,
        DigitCount := HexDigitCount);
    Message := CONCAT('Assertion failed: bit value does not match. BitIndex = ',
        USINT_TO_STRING(BitIndex));
    Message := CONCAT(Message, ', Expected = ');
    Message := CONCAT(Message, BOOL_TO_STRING(Expected));
    Message := CONCAT(Message, ', Actual = ');
    Message := CONCAT(Message, BOOL_TO_STRING(ActualBit));
    Message := CONCAT(Message, ', Value = ');
    Message := CONCAT(Message, ActualText);
    Message := CONCAT(Message, '.');
    Fail(Message := Message);
    RETURN;
END_IF;

Pass();
END_METHOD

END_FUNCTION_BLOCK

// ---- Framework/Assertions/POU/BasicTypes/LWord/AssertEqualMask_LWord.TcPOU
{region 'Documentation'}
(*!
<summary>Checks that selected bits match the expected masked value.</summary>
*)
{endregion}
FUNCTION_BLOCK AssertEqualMask_LWord EXTENDS AssertionBase
VAR_INPUT
    IN : LWORD; //! Actual bitfield.
    Mask : LWORD := 16#FFFFFFFFFFFFFFFF; //! Selects evaluated bits; defaults to all bits. An empty mask produces Error during evaluation.
    Expected : LWORD; //! Expected value; bits outside Mask are ignored.
END_VAR

SUPER^();

{region 'Documentation'}
(*!
<summary>Rejects an empty mask before comparing selected bits.</summary>
*)
{endregion}
METHOD PROTECTED Assert
VAR
    Message : STRING(GVL_Constants.MessageLength);
    MaskText : STRING(GVL_Constants.AssertionValueLength);
    ExpectedText : STRING(GVL_Constants.AssertionValueLength);
    ActualText : STRING(GVL_Constants.AssertionValueLength);
END_VAR
VAR CONSTANT
    NoMask : LWORD := 16#00;
    HexDigitCount : USINT := 16;
END_VAR
IF NOT EvaluationActive THEN
    RETURN;
END_IF;

IF Result = E_Result.Error THEN
    RETURN;
END_IF;

IF Mask = NoMask THEN
    MaskText := CreateAssertionTextValue_Hex(Value := Mask,
        DigitCount := HexDigitCount);
    Message := CONCAT('Assertion error: mask must not be empty. Mask = ',
        MaskText);
    Message := CONCAT(Message, '.');
    Error(Message := Message);
    RETURN;
END_IF;

IF Result = E_Result.Failed THEN
    RETURN;
END_IF;

IF (IN AND Mask) <> (Expected AND Mask) THEN
    MaskText := CreateAssertionTextValue_Hex(Value := Mask,
        DigitCount := HexDigitCount);
    ExpectedText := CreateAssertionTextValue_Hex(Value := Expected,
        DigitCount := HexDigitCount);
    ActualText := CreateAssertionTextValue_Hex(Value := IN,
        DigitCount := HexDigitCount);
    Message := CONCAT('Assertion failed: selected bits do not match. Expected = ',
        ExpectedText);
    Message := CONCAT(Message, ', Mask = ');
    Message := CONCAT(Message, MaskText);
    Message := CONCAT(Message, ', Actual = ');
    Message := CONCAT(Message, ActualText);
    Message := CONCAT(Message, '.');
    Fail(Message := Message);
    RETURN;
END_IF;

Pass();
END_METHOD

END_FUNCTION_BLOCK

// ---- Framework/Assertions/POU/BasicTypes/LWord/AssertFalseBit_LWord.TcPOU
{region 'Documentation'}
(*!
<summary>Checks that the selected LWORD bit is FALSE.</summary>
*)
{endregion}
FUNCTION_BLOCK AssertFalseBit_LWord EXTENDS AssertionBase
VAR_INPUT
    IN : LWORD; //! Actual bitfield.
    BitIndex : USINT; //! Zero-based bit index (0..63); an invalid index produces Error during evaluation.
END_VAR

SUPER^();

{region 'Documentation'}
(*!
<summary>Validates the index before evaluating the selected bit.</summary>
*)
{endregion}
METHOD PROTECTED Assert
VAR
    Mask : LWORD;
    ActualBit : BOOL;
    Message : STRING(GVL_Constants.MessageLength);
    ActualText : STRING(GVL_Constants.AssertionValueLength);
END_VAR
VAR CONSTANT
    MaxBitIndex : USINT := 63;
    SingleBitMask : LWORD := 16#01;
    NoBitMask : LWORD := 16#00;
    HexDigitCount : USINT := 16;
END_VAR
IF NOT EvaluationActive THEN
    RETURN;
END_IF;

IF Result = E_Result.Error THEN
    RETURN;
END_IF;

IF BitIndex > MaxBitIndex THEN
    Message := CONCAT('Assertion error: bit index is outside valid range. BitIndex = ',
        USINT_TO_STRING(BitIndex));
    Message := CONCAT(Message, ', MaxBitIndex = ');
    Message := CONCAT(Message, USINT_TO_STRING(MaxBitIndex));
    Message := CONCAT(Message, '.');
    Error(Message := Message);
    RETURN;
END_IF;

IF Result = E_Result.Failed THEN
    RETURN;
END_IF;

Mask := SHL(SingleBitMask, BitIndex);
ActualBit := (IN AND Mask) <> NoBitMask;

IF ActualBit THEN
    ActualText := CreateAssertionTextValue_Hex(Value := IN,
        DigitCount := HexDigitCount);
    Message := CONCAT('Assertion failed: bit is TRUE but must be FALSE. BitIndex = ',
        USINT_TO_STRING(BitIndex));
    Message := CONCAT(Message, ', Actual = ');
    Message := CONCAT(Message, ActualText);
    Message := CONCAT(Message, '.');
    Fail(Message := Message);
    RETURN;
END_IF;

Pass();
END_METHOD

END_FUNCTION_BLOCK

// ---- Framework/Assertions/POU/BasicTypes/LWord/AssertFalseMask_LWord.TcPOU
{region 'Documentation'}
(*!
<summary>Checks that all selected bits are FALSE.</summary>
*)
{endregion}
FUNCTION_BLOCK AssertFalseMask_LWord EXTENDS AssertionBase
VAR_INPUT
    IN : LWORD; //! Actual bitfield.
    Mask : LWORD := 16#FFFFFFFFFFFFFFFF; //! Selects evaluated bits; defaults to all bits. An empty mask produces Error during evaluation.
END_VAR

SUPER^();

{region 'Documentation'}
(*!
<summary>Rejects an empty mask before comparing selected bits.</summary>
*)
{endregion}
METHOD PROTECTED Assert
VAR
    Message : STRING(GVL_Constants.MessageLength);
    MaskText : STRING(GVL_Constants.AssertionValueLength);
    ActualText : STRING(GVL_Constants.AssertionValueLength);
END_VAR
VAR CONSTANT
    NoMask : LWORD := 16#00;
    HexDigitCount : USINT := 16;
END_VAR
IF NOT EvaluationActive THEN
    RETURN;
END_IF;

IF Result = E_Result.Error THEN
    RETURN;
END_IF;

IF Mask = NoMask THEN
    MaskText := CreateAssertionTextValue_Hex(Value := Mask,
        DigitCount := HexDigitCount);
    Message := CONCAT('Assertion error: mask must not be empty. Mask = ',
        MaskText);
    Message := CONCAT(Message, '.');
    Error(Message := Message);
    RETURN;
END_IF;

IF Result = E_Result.Failed THEN
    RETURN;
END_IF;

IF (IN AND Mask) <> NoMask THEN
    MaskText := CreateAssertionTextValue_Hex(Value := Mask,
        DigitCount := HexDigitCount);
    ActualText := CreateAssertionTextValue_Hex(Value := IN,
        DigitCount := HexDigitCount);
    Message := CONCAT('Assertion failed: selected bits are not all FALSE. Mask = ',
        MaskText);
    Message := CONCAT(Message, ', Actual = ');
    Message := CONCAT(Message, ActualText);
    Message := CONCAT(Message, '.');
    Fail(Message := Message);
    RETURN;
END_IF;

Pass();
END_METHOD

END_FUNCTION_BLOCK

// ---- Framework/Assertions/POU/BasicTypes/LWord/AssertNotEqualBit_LWord.TcPOU
{region 'Documentation'}
(*!
<summary>Checks that the selected LWORD bit differs from the expected Boolean value.</summary>
*)
{endregion}
FUNCTION_BLOCK AssertNotEqualBit_LWord EXTENDS AssertionBase
VAR_INPUT
    IN : LWORD; //! Actual bitfield.
    BitIndex : USINT; //! Zero-based bit index (0..63); an invalid index produces Error during evaluation.
    Expected : BOOL; //! Forbidden selected bit value.
END_VAR

SUPER^();

{region 'Documentation'}
(*!
<summary>Validates the index before evaluating the selected bit.</summary>
*)
{endregion}
METHOD PROTECTED Assert
VAR
    Mask : LWORD;
    ActualBit : BOOL;
    Message : STRING(GVL_Constants.MessageLength);
    ActualText : STRING(GVL_Constants.AssertionValueLength);
END_VAR
VAR CONSTANT
    MaxBitIndex : USINT := 63;
    SingleBitMask : LWORD := 16#01;
    NoBitMask : LWORD := 16#00;
    HexDigitCount : USINT := 16;
END_VAR
IF NOT EvaluationActive THEN
    RETURN;
END_IF;

IF Result = E_Result.Error THEN
    RETURN;
END_IF;

IF BitIndex > MaxBitIndex THEN
    Message := CONCAT('Assertion error: bit index is outside valid range. BitIndex = ',
        USINT_TO_STRING(BitIndex));
    Message := CONCAT(Message, ', MaxBitIndex = ');
    Message := CONCAT(Message, USINT_TO_STRING(MaxBitIndex));
    Message := CONCAT(Message, '.');
    Error(Message := Message);
    RETURN;
END_IF;

IF Result = E_Result.Failed THEN
    RETURN;
END_IF;

Mask := SHL(SingleBitMask, BitIndex);
ActualBit := (IN AND Mask) <> NoBitMask;

IF ActualBit = Expected THEN
    ActualText := CreateAssertionTextValue_Hex(Value := IN,
        DigitCount := HexDigitCount);
    Message := CONCAT('Assertion failed: bit value matches forbidden value. BitIndex = ',
        USINT_TO_STRING(BitIndex));
    Message := CONCAT(Message, ', NotExpected = ');
    Message := CONCAT(Message, BOOL_TO_STRING(Expected));
    Message := CONCAT(Message, ', Actual = ');
    Message := CONCAT(Message, BOOL_TO_STRING(ActualBit));
    Message := CONCAT(Message, ', Value = ');
    Message := CONCAT(Message, ActualText);
    Message := CONCAT(Message, '.');
    Fail(Message := Message);
    RETURN;
END_IF;

Pass();
END_METHOD

END_FUNCTION_BLOCK

// ---- Framework/Assertions/POU/BasicTypes/LWord/AssertNoValueChange_LWord.TcPOU
{region 'Documentation'}
(*!
<summary>Check equality between consecutive active observations.</summary>
<description>

The first active observation establishes a baseline without deciding a result. Disabling
observation invalidates that baseline, not the held Result. Re-enabling first establishes a new
baseline; Reset clears history.

ObserveFirstCycle FALSE delays the first observation by one enabled call.

</description>
*)
{endregion}
FUNCTION_BLOCK AssertNoValueChange_LWord EXTENDS AssertionBase
VAR_INPUT
    IN : LWORD; //! Actual value to observe.
END_VAR
VAR
    FINPrevious : LWORD;
    FObservationPrevious : BOOL;
    FEvaluationActive : BOOL;
END_VAR

SUPER^();

{region 'Documentation'}
(*!
<summary>Observe the current value before evaluating a change against the previous observation.</summary>
*)
{endregion}
METHOD PROTECTED Assert
VAR
    PreviousValue : LWORD;
    Message : STRING(GVL_Constants.MessageLength);
    PreviousText : STRING(GVL_Constants.AssertionValueLength);
    ActualText : STRING(GVL_Constants.AssertionValueLength);
END_VAR
VAR CONSTANT
    HexDigitCount : USINT := 16;
END_VAR
FEvaluationActive := ObservationActive AND FObservationPrevious;
FObservationPrevious := ObservationActive;

IF NOT ObservationActive THEN
    RETURN;
END_IF;

PreviousValue := FINPrevious;
FINPrevious := IN;

IF NOT EvaluationActive THEN
    RETURN;
END_IF;

IF Result = E_Result.Error THEN
    RETURN;
END_IF;

IF Result = E_Result.Failed THEN
    RETURN;
END_IF;

IF IN <> PreviousValue THEN
    PreviousText := CreateAssertionTextValue_Hex(Value := PreviousValue,
        DigitCount := HexDigitCount);
    ActualText := CreateAssertionTextValue_Hex(Value := IN,
        DigitCount := HexDigitCount);
    Message := CONCAT('Assertion failed: value changed unexpectedly. Previous = ',
        PreviousText);
    Message := CONCAT(Message, ', Actual = ');
    Message := CONCAT(Message, ActualText);
    Message := CONCAT(Message, '.');
    Fail(Message := Message);
    RETURN;
END_IF;

Pass();
END_METHOD

{region 'Documentation'}
(*!
<summary>Current/last call has an active observation and a preceding observation
baseline.</summary>
*)
{endregion}
{attribute 'monitoring' := 'call'}
PROPERTY PUBLIC EvaluationActive : BOOL //! Current/last call has an active observation and a preceding observation baseline.
GET // PUBLIC
EvaluationActive := FEvaluationActive;
END_GET
END_PROPERTY

{region 'Documentation'}
(*!
<summary>Clear observation history and the current evaluation gate.</summary>
*)
{endregion}
METHOD PROTECTED ResetAssertion
FINPrevious := 0;
FObservationPrevious := FALSE;
FEvaluationActive := FALSE;
END_METHOD

END_FUNCTION_BLOCK

// ---- Framework/Assertions/POU/AssertionEdgeCountBase.TcPOU
{region 'Documentation'}
(*!
<summary>Shared edge observation and bounded cumulative count for explicit-evaluation
assertions.</summary>
<description>

Derived Assert implementations call SUPER^.Assert() once before evaluating the count.
Implement the side-effect-free IsMatchingEdge predicate for rising or falling edges.

The first active observation establishes a signal baseline without counting an edge. An
observation interruption invalidates that baseline but retains the accumulated count until
Reset. Evaluate checks that count independently of Enable.

The UINT count saturates at 65535. The next matching edge reports Error rather than
wrapping; this observation error can occur without explicit evaluation.

</description>
*)
{endregion}
FUNCTION_BLOCK ABSTRACT AssertionEdgeCountBase EXTENDS AssertionWithEvaluationBase
VAR_INPUT
    IN : BOOL; //! Signal sampled while ObservationActive; the first sample establishes the edge baseline.
END_VAR
VAR
    FINPrevious : BOOL;
    FObservationPrevious : BOOL;
    FEdgeCount : UINT;
END_VAR
VAR CONSTANT
    MaxEdgeCount : UINT := 65535;
END_VAR

SUPER^();

{region 'Documentation'}
(*!
<summary>Capture history and count a matching edge before independent result
evaluation.</summary>
*)
{endregion}
METHOD PROTECTED Assert
VAR
    HasPreviousObservation : BOOL;
    PreviousValue : BOOL;
END_VAR
HasPreviousObservation := FObservationPrevious;
FObservationPrevious := ObservationActive;

IF NOT ObservationActive THEN
    RETURN;
END_IF;

PreviousValue := FINPrevious;
FINPrevious := IN;

IF NOT HasPreviousObservation THEN
    RETURN;
END_IF;

IF NOT IsMatchingEdge(PreviousValue := PreviousValue,
    CurrentValue := IN) THEN
    RETURN;
END_IF;

IF FEdgeCount = MaxEdgeCount THEN
    Error(Message := 'Assertion error: edge count exceeds UINT capacity.');
    RETURN;
END_IF;

FEdgeCount := FEdgeCount + 1;
END_METHOD

{region 'Documentation'}
(*!
<summary>Observed edges; retained across observation interruptions and cleared by
Reset.</summary>
*)
{endregion}
{attribute 'monitoring' := 'call'}
PROPERTY PUBLIC EdgeCount : UINT //! Observed edges; retained across observation interruptions and cleared by Reset.
GET // PUBLIC
EdgeCount := FEdgeCount;
END_GET
END_PROPERTY

{region 'Documentation'}
(*!
<summary>Return whether the two observed values form the selected edge; no side
effects.</summary>
*)
{endregion}
METHOD PROTECTED ABSTRACT IsMatchingEdge : BOOL //! TRUE when PreviousValue and CurrentValue form the edge selected by this Assertion.
VAR_INPUT
    PreviousValue : BOOL; //! Signal value from the preceding active observation.
    CurrentValue : BOOL; //! Signal value from the current active observation.
END_VAR
END_METHOD

{region 'Documentation'}
(*!
<summary>Clear edge count and invalidate the observation baseline.</summary>
*)
{endregion}
METHOD PROTECTED ResetAssertion
FINPrevious := FALSE;
FObservationPrevious := FALSE;
FEdgeCount := 0;
END_METHOD

END_FUNCTION_BLOCK

// ---- Framework/Assertions/POU/Utilities/CountArrayTokens_Byte.TcPOU
{region 'Documentation'}
(*!
<summary>Counts exact non-overlapping tokens; advances past each complete match. Caller validates stable references, a nonempty in-bounds range and a nonempty token fitting the range.</summary>
*)
{endregion}
FUNCTION INTERNAL CountArrayTokens_Byte : UINT //! Number of non-overlapping token occurrences in the selected range.
VAR_INPUT
    StartIndex : DINT; //! First selected index in IN; uses the array's declared index range, not a zero-based offset.
    Length : USINT; //! Number of selected elements starting at StartIndex; must fit the array range; valid range 1..255.
END_VAR
VAR_IN_OUT CONSTANT
    IN : ARRAY[*] OF BYTE; //! Read-only actual data; the selected range must remain stable during the call.
    Token : ARRAY[*] OF BYTE; //! Read-only nonempty token; keep stable during the call and within the selected search length.
END_VAR
VAR
    CandidateOffset : LINT;
    LastCandidateOffset : LINT;
    TokenLowerIndex : DINT;
    TokenLength : LINT;
    TokenOffset : LINT;
    InIndex : DINT;
    TokenIndex : DINT;
    TokenMatches : BOOL;
END_VAR

CountArrayTokens_Byte := 0;
TokenLowerIndex := LOWER_BOUND(Token, 1);
TokenLength := DINT_TO_LINT(UPPER_BOUND(Token, 1)) - DINT_TO_LINT(TokenLowerIndex) + 1;
LastCandidateOffset := USINT_TO_LINT(Length) - TokenLength;
CandidateOffset := 0;

WHILE CandidateOffset <= LastCandidateOffset DO
    TokenMatches := TRUE;
    FOR TokenOffset := 0 TO TokenLength - 1 DO
        InIndex := LINT_TO_DINT(DINT_TO_LINT(StartIndex) + CandidateOffset + TokenOffset);
        TokenIndex := LINT_TO_DINT(DINT_TO_LINT(TokenLowerIndex) + TokenOffset);
        IF IN[InIndex] <> Token[TokenIndex] THEN
            TokenMatches := FALSE;
            EXIT;
        END_IF;
    END_FOR;

    IF TokenMatches THEN
        CountArrayTokens_Byte := CountArrayTokens_Byte + 1;
        CandidateOffset := CandidateOffset + TokenLength;
    ELSE
        CandidateOffset := CandidateOffset + 1;
    END_IF;
END_WHILE;

END_FUNCTION

// ---- Framework/Assertions/POU/Utilities/CountArrayTokens_Word.TcPOU
{region 'Documentation'}
(*!
<summary>Counts exact non-overlapping tokens; advances past each complete match. Caller validates stable references, a nonempty in-bounds range and a nonempty token fitting the range.</summary>
*)
{endregion}
FUNCTION INTERNAL CountArrayTokens_Word : UINT //! Number of non-overlapping token occurrences in the selected range.
VAR_INPUT
    StartIndex : DINT; //! First selected index in IN; uses the array's declared index range, not a zero-based offset.
    Length : USINT; //! Number of selected elements starting at StartIndex; must fit the array range; valid range 1..255.
END_VAR
VAR_IN_OUT CONSTANT
    IN : ARRAY[*] OF WORD; //! Read-only actual data; the selected range must remain stable during the call.
    Token : ARRAY[*] OF WORD; //! Read-only nonempty token; keep stable during the call and within the selected search length.
END_VAR
VAR
    CandidateOffset : LINT;
    LastCandidateOffset : LINT;
    TokenLowerIndex : DINT;
    TokenLength : LINT;
    TokenOffset : LINT;
    InIndex : DINT;
    TokenIndex : DINT;
    TokenMatches : BOOL;
END_VAR

CountArrayTokens_Word := 0;
TokenLowerIndex := LOWER_BOUND(Token, 1);
TokenLength := DINT_TO_LINT(UPPER_BOUND(Token, 1)) - DINT_TO_LINT(TokenLowerIndex) + 1;
LastCandidateOffset := USINT_TO_LINT(Length) - TokenLength;
CandidateOffset := 0;

WHILE CandidateOffset <= LastCandidateOffset DO
    TokenMatches := TRUE;
    FOR TokenOffset := 0 TO TokenLength - 1 DO
        InIndex := LINT_TO_DINT(DINT_TO_LINT(StartIndex) + CandidateOffset + TokenOffset);
        TokenIndex := LINT_TO_DINT(DINT_TO_LINT(TokenLowerIndex) + TokenOffset);
        IF IN[InIndex] <> Token[TokenIndex] THEN
            TokenMatches := FALSE;
            EXIT;
        END_IF;
    END_FOR;

    IF TokenMatches THEN
        CountArrayTokens_Word := CountArrayTokens_Word + 1;
        CandidateOffset := CandidateOffset + TokenLength;
    ELSE
        CandidateOffset := CandidateOffset + 1;
    END_IF;
END_WHILE;

END_FUNCTION

// ---- Framework/Assertions/POU/Utilities/CountValueTokens_Byte.TcPOU
{region 'Documentation'}
(*!
<summary>Counts all masked value matches in the selected range. Caller validates stable references, a nonempty in-bounds range.</summary>
*)
{endregion}
FUNCTION INTERNAL CountValueTokens_Byte : UINT //! Number of masked value matches in the selected range.
VAR_INPUT
    StartIndex : DINT; //! First selected index in IN; uses the array's declared index range, not a zero-based offset.
    Length : USINT; //! Number of selected elements starting at StartIndex; must fit the array range; valid range 1..255.
    Token : BYTE; //! Value searched for in the selected range; Mask selects the compared bits.
    Mask : BYTE; //! Bits included in the comparison; bits outside the mask are ignored.
END_VAR
VAR_IN_OUT CONSTANT
    IN : ARRAY[*] OF BYTE; //! Read-only actual data; the selected range must remain stable during the call.
END_VAR
VAR
    CandidateOffset : LINT;
    InIndex : DINT;
END_VAR

CountValueTokens_Byte := 0;

FOR CandidateOffset := 0 TO USINT_TO_LINT(Length) - 1 DO
    InIndex := LINT_TO_DINT(DINT_TO_LINT(StartIndex) + CandidateOffset);
    IF (IN[InIndex] AND Mask) = (Token AND Mask) THEN
        CountValueTokens_Byte := CountValueTokens_Byte + 1;
    END_IF;
END_FOR;

END_FUNCTION

// ---- Framework/Assertions/POU/Utilities/CountValueTokens_Word.TcPOU
{region 'Documentation'}
(*!
<summary>Counts all masked value matches in the selected range. Caller validates stable references, a nonempty in-bounds range.</summary>
*)
{endregion}
FUNCTION INTERNAL CountValueTokens_Word : UINT //! Number of masked value matches in the selected range.
VAR_INPUT
    StartIndex : DINT; //! First selected index in IN; uses the array's declared index range, not a zero-based offset.
    Length : USINT; //! Number of selected elements starting at StartIndex; must fit the array range; valid range 1..255.
    Token : WORD; //! Value searched for in the selected range; Mask selects the compared bits.
    Mask : WORD; //! Bits included in the comparison; bits outside the mask are ignored.
END_VAR
VAR_IN_OUT CONSTANT
    IN : ARRAY[*] OF WORD; //! Read-only actual data; the selected range must remain stable during the call.
END_VAR
VAR
    CandidateOffset : LINT;
    InIndex : DINT;
END_VAR

CountValueTokens_Word := 0;

FOR CandidateOffset := 0 TO USINT_TO_LINT(Length) - 1 DO
    InIndex := LINT_TO_DINT(DINT_TO_LINT(StartIndex) + CandidateOffset);
    IF (IN[InIndex] AND Mask) = (Token AND Mask) THEN
        CountValueTokens_Word := CountValueTokens_Word + 1;
    END_IF;
END_FOR;

END_FUNCTION

// ---- Framework/Assertions/POU/Utilities/FindArrayToken_Byte.TcPOU
{region 'Documentation'}
(*!
<summary>Finds the first exact contiguous array token in the selected range. Caller validates stable references, a nonempty in-bounds range, and a nonempty token fitting the range.</summary>
*)
{endregion}
FUNCTION INTERNAL FindArrayToken_Byte : BOOL //! TRUE when a token was found; Index is its absolute array index and may legitimately be zero.
VAR_INPUT
    StartIndex : DINT; //! First selected index in IN; uses the array's declared index range, not a zero-based offset.
    Length : USINT; //! Number of selected elements starting at StartIndex; must fit the array range; valid range 1..255.
END_VAR
VAR_OUTPUT
    Index : DINT; //! Absolute matching index; zero when no match exists. Use the BOOL result to distinguish.
END_VAR
VAR_IN_OUT CONSTANT
    IN : ARRAY[*] OF BYTE; //! Read-only actual data; the selected range must remain stable during the call.
    Token : ARRAY[*] OF BYTE; //! Read-only nonempty token; keep stable during the call and within the selected search length.
END_VAR
VAR
    CandidateOffset : LINT;
    InIndex : DINT;
    TokenLowerIndex : DINT;
    TokenLength : LINT;
    TokenOffset : LINT;
    TokenIndex : DINT;
    TokenMatches : BOOL;
END_VAR

FindArrayToken_Byte := FALSE;
Index := 0;

TokenLowerIndex := LOWER_BOUND(Token, 1);
TokenLength := DINT_TO_LINT(UPPER_BOUND(Token, 1)) - DINT_TO_LINT(TokenLowerIndex) + 1;

FOR CandidateOffset := 0 TO USINT_TO_LINT(Length) - TokenLength DO
    TokenMatches := TRUE;
    FOR TokenOffset := 0 TO TokenLength - 1 DO
        InIndex := LINT_TO_DINT(DINT_TO_LINT(StartIndex) + CandidateOffset + TokenOffset);
        TokenIndex := LINT_TO_DINT(DINT_TO_LINT(TokenLowerIndex) + TokenOffset);
        IF IN[InIndex] <> Token[TokenIndex] THEN
            TokenMatches := FALSE;
            EXIT;
        END_IF;
    END_FOR;
    IF TokenMatches THEN
        Index := LINT_TO_DINT(DINT_TO_LINT(StartIndex) + CandidateOffset);
        FindArrayToken_Byte := TRUE;
        RETURN;
    END_IF;
END_FOR;

END_FUNCTION

// ---- Framework/Assertions/POU/Utilities/FindArrayToken_Word.TcPOU
{region 'Documentation'}
(*!
<summary>Finds the first exact contiguous array token in the selected range. Caller validates stable references, a nonempty in-bounds range, and a nonempty token fitting the range.</summary>
*)
{endregion}
FUNCTION INTERNAL FindArrayToken_Word : BOOL //! TRUE when a token was found; Index is its absolute array index and may legitimately be zero.
VAR_INPUT
    StartIndex : DINT; //! First selected index in IN; uses the array's declared index range, not a zero-based offset.
    Length : USINT; //! Number of selected elements starting at StartIndex; must fit the array range; valid range 1..255.
END_VAR
VAR_OUTPUT
    Index : DINT; //! Absolute matching index; zero when no match exists. Use the BOOL result to distinguish.
END_VAR
VAR_IN_OUT CONSTANT
    IN : ARRAY[*] OF WORD; //! Read-only actual data; the selected range must remain stable during the call.
    Token : ARRAY[*] OF WORD; //! Read-only nonempty token; keep stable during the call and within the selected search length.
END_VAR
VAR
    CandidateOffset : LINT;
    InIndex : DINT;
    TokenLowerIndex : DINT;
    TokenLength : LINT;
    TokenOffset : LINT;
    TokenIndex : DINT;
    TokenMatches : BOOL;
END_VAR

FindArrayToken_Word := FALSE;
Index := 0;

TokenLowerIndex := LOWER_BOUND(Token, 1);
TokenLength := DINT_TO_LINT(UPPER_BOUND(Token, 1)) - DINT_TO_LINT(TokenLowerIndex) + 1;

FOR CandidateOffset := 0 TO USINT_TO_LINT(Length) - TokenLength DO
    TokenMatches := TRUE;
    FOR TokenOffset := 0 TO TokenLength - 1 DO
        InIndex := LINT_TO_DINT(DINT_TO_LINT(StartIndex) + CandidateOffset + TokenOffset);
        TokenIndex := LINT_TO_DINT(DINT_TO_LINT(TokenLowerIndex) + TokenOffset);
        IF IN[InIndex] <> Token[TokenIndex] THEN
            TokenMatches := FALSE;
            EXIT;
        END_IF;
    END_FOR;
    IF TokenMatches THEN
        Index := LINT_TO_DINT(DINT_TO_LINT(StartIndex) + CandidateOffset);
        FindArrayToken_Word := TRUE;
        RETURN;
    END_IF;
END_FOR;

END_FUNCTION

// ---- Framework/Assertions/POU/Utilities/FindValueToken_Byte.TcPOU
{region 'Documentation'}
(*!
<summary>Finds the first masked value token in the selected range. Caller validates stable references, a nonempty in-bounds range.</summary>
*)
{endregion}
FUNCTION INTERNAL FindValueToken_Byte : BOOL //! TRUE when a token was found; Index is its absolute array index and may legitimately be zero.
VAR_INPUT
    StartIndex : DINT; //! First selected index in IN; uses the array's declared index range, not a zero-based offset.
    Length : USINT; //! Number of selected elements starting at StartIndex; must fit the array range; valid range 1..255.
    Token : BYTE; //! Value searched for in the selected range; Mask selects the compared bits.
    Mask : BYTE; //! Bits included in the comparison; bits outside the mask are ignored.
END_VAR
VAR_OUTPUT
    Index : DINT; //! Absolute matching index; zero when no match exists. Use the BOOL result to distinguish.
END_VAR
VAR_IN_OUT CONSTANT
    IN : ARRAY[*] OF BYTE; //! Read-only actual data; the selected range must remain stable during the call.
END_VAR
VAR
    CandidateOffset : LINT;
    InIndex : DINT;
END_VAR

FindValueToken_Byte := FALSE;
Index := 0;

FOR CandidateOffset := 0 TO USINT_TO_LINT(Length) - 1 DO
    InIndex := LINT_TO_DINT(DINT_TO_LINT(StartIndex) + CandidateOffset);
    IF (IN[InIndex] AND Mask) = (Token AND Mask) THEN
        Index := LINT_TO_DINT(DINT_TO_LINT(StartIndex) + CandidateOffset);
        FindValueToken_Byte := TRUE;
        RETURN;
    END_IF;
END_FOR;

END_FUNCTION

// ---- Framework/Assertions/POU/Utilities/FindValueToken_Word.TcPOU
{region 'Documentation'}
(*!
<summary>Finds the first masked value token in the selected range. Caller validates stable references, a nonempty in-bounds range.</summary>
*)
{endregion}
FUNCTION INTERNAL FindValueToken_Word : BOOL //! TRUE when a token was found; Index is its absolute array index and may legitimately be zero.
VAR_INPUT
    StartIndex : DINT; //! First selected index in IN; uses the array's declared index range, not a zero-based offset.
    Length : USINT; //! Number of selected elements starting at StartIndex; must fit the array range; valid range 1..255.
    Token : WORD; //! Value searched for in the selected range; Mask selects the compared bits.
    Mask : WORD; //! Bits included in the comparison; bits outside the mask are ignored.
END_VAR
VAR_OUTPUT
    Index : DINT; //! Absolute matching index; zero when no match exists. Use the BOOL result to distinguish.
END_VAR
VAR_IN_OUT CONSTANT
    IN : ARRAY[*] OF WORD; //! Read-only actual data; the selected range must remain stable during the call.
END_VAR
VAR
    CandidateOffset : LINT;
    InIndex : DINT;
END_VAR

FindValueToken_Word := FALSE;
Index := 0;

FOR CandidateOffset := 0 TO USINT_TO_LINT(Length) - 1 DO
    InIndex := LINT_TO_DINT(DINT_TO_LINT(StartIndex) + CandidateOffset);
    IF (IN[InIndex] AND Mask) = (Token AND Mask) THEN
        Index := LINT_TO_DINT(DINT_TO_LINT(StartIndex) + CandidateOffset);
        FindValueToken_Word := TRUE;
        RETURN;
    END_IF;
END_FOR;

END_FUNCTION

// ---- Framework/Assertions/POU/Utilities/IsTimeOfDayValid_TOD.TcPOU
{region 'Documentation'}
(*!
<summary>Checks the native time-of-day range without changing or normalizing Value.</summary>
*)
{endregion}
FUNCTION INTERNAL IsTimeOfDayValid_TOD : BOOL //! TRUE for a time of day below 24 hours; the value is not normalized.
VAR_INPUT
    Value : TOD; //! Time-of-day value checked against the interval from midnight inclusive to the next midnight exclusive.
END_VAR
VAR CONSTANT
    MaximumTimeOfDay : TOD := TOD#23:59:59.999;
END_VAR

IsTimeOfDayValid_TOD := Value <= MaximumTimeOfDay;

END_FUNCTION

// ---- Framework/Assertions/POU/Utilities/TextContains_String.TcPOU
{region 'Documentation'}
(*!
<summary>Searches for a nonempty fragment by exact code-unit comparison without copies. Caller supplies valid, stable references and content within the configured assertion capacity.</summary>
*)
{endregion}
FUNCTION INTERNAL TextContains_String : BOOL //! TRUE when the nonempty Fragment occurs in Value.
VAR_IN_OUT CONSTANT
    Value : STRING(Param_Assertions.AssertionStringLength); //! Read-only source text; must be terminated within the configured capacity and stable during the call.
    Fragment : STRING(Param_Assertions.AssertionStringLength); //! Read-only nonempty text fragment searched for in Value.
END_VAR
VAR
    ValueLength : DINT;
    FragmentLength : DINT;
    StartIndex : DINT;
    CharacterIndex : DINT;
    MatchesFragment : BOOL;
END_VAR
VAR CONSTANT
    Terminator : BYTE := 0;
END_VAR

TextContains_String := FALSE;

FOR ValueLength := 0 TO UINT_TO_DINT(Param_Assertions.AssertionStringLength) DO
    // SA0175: Exact byte comparison; caller validates termination/capacity and indices stay in bounds.
    {analysis -175}
    IF Value[ValueLength] = Terminator THEN
    {analysis +175}
        EXIT;
    END_IF;
END_FOR;

FOR FragmentLength := 0 TO UINT_TO_DINT(Param_Assertions.AssertionStringLength) DO
    // SA0175: Exact byte comparison; caller validates termination/capacity and indices stay in bounds.
    {analysis -175}
    IF Fragment[FragmentLength] = Terminator THEN
    {analysis +175}
        EXIT;
    END_IF;
END_FOR;

IF (FragmentLength = 0) OR (FragmentLength > ValueLength) THEN
    RETURN;
END_IF;

FOR StartIndex := 0 TO ValueLength - FragmentLength DO
    MatchesFragment := TRUE;
    FOR CharacterIndex := 0 TO FragmentLength - 1 DO
        // SA0175: Exact byte comparison; caller validates termination/capacity and indices stay in bounds.
        {analysis -175}
        IF Value[StartIndex + CharacterIndex] <> Fragment[CharacterIndex] THEN
        {analysis +175}
            MatchesFragment := FALSE;
            EXIT;
        END_IF;
    END_FOR;

    IF MatchesFragment THEN
        TextContains_String := TRUE;
        RETURN;
    END_IF;
END_FOR;

END_FUNCTION

// ---- Framework/Assertions/POU/Utilities/TextContains_WString.TcPOU
{region 'Documentation'}
(*!
<summary>Searches for a nonempty fragment by exact code-unit comparison without copies. Caller supplies valid, stable references and content within the configured assertion capacity.</summary>
*)
{endregion}
FUNCTION INTERNAL TextContains_WString : BOOL //! TRUE when the nonempty Fragment occurs in Value.
VAR_IN_OUT CONSTANT
    Value : WSTRING(Param_Assertions.AssertionWStringLength); //! Read-only source text; must be terminated within the configured capacity and stable during the call.
    Fragment : WSTRING(Param_Assertions.AssertionWStringLength); //! Read-only nonempty text fragment searched for in Value.
END_VAR
VAR
    ValueLength : DINT;
    FragmentLength : DINT;
    StartIndex : DINT;
    CharacterIndex : DINT;
    MatchesFragment : BOOL;
END_VAR
VAR CONSTANT
    Terminator : WORD := 0;
END_VAR

TextContains_WString := FALSE;

FOR ValueLength := 0 TO UINT_TO_DINT(Param_Assertions.AssertionWStringLength) DO
    IF Value[ValueLength] = Terminator THEN
        EXIT;
    END_IF;
END_FOR;

FOR FragmentLength := 0 TO UINT_TO_DINT(Param_Assertions.AssertionWStringLength) DO
    IF Fragment[FragmentLength] = Terminator THEN
        EXIT;
    END_IF;
END_FOR;

IF (FragmentLength = 0) OR (FragmentLength > ValueLength) THEN
    RETURN;
END_IF;

FOR StartIndex := 0 TO ValueLength - FragmentLength DO
    MatchesFragment := TRUE;
    FOR CharacterIndex := 0 TO FragmentLength - 1 DO
        IF Value[StartIndex + CharacterIndex] <> Fragment[CharacterIndex] THEN
            MatchesFragment := FALSE;
            EXIT;
        END_IF;
    END_FOR;

    IF MatchesFragment THEN
        TextContains_WString := TRUE;
        RETURN;
    END_IF;
END_FOR;

END_FUNCTION

// ---- Framework/Assertions/POU/Utilities/TextEndsWith_String.TcPOU
{region 'Documentation'}
(*!
<summary>Exact suffix comparison without copies; an empty suffix matches. Caller supplies valid, stable references and content within the configured assertion capacity.</summary>
*)
{endregion}
FUNCTION INTERNAL TextEndsWith_String : BOOL //! TRUE when Value ends with Suffix; an empty Suffix matches.
VAR_IN_OUT CONSTANT
    Value : STRING(Param_Assertions.AssertionStringLength); //! Read-only source text; must be terminated within the configured capacity and stable during the call.
    Suffix : STRING(Param_Assertions.AssertionStringLength); //! Read-only suffix compared by code unit; an empty value matches in this helper.
END_VAR
VAR
    CharacterIndex : DINT;
    ValueLength : DINT;
    SuffixLength : DINT;
    SuffixStartIndex : DINT;
END_VAR
VAR CONSTANT
    Terminator : BYTE := 0;
END_VAR

TextEndsWith_String := FALSE;

FOR ValueLength := 0 TO UINT_TO_DINT(Param_Assertions.AssertionStringLength) DO
    // SA0175: Exact byte comparison; caller validates termination/capacity and indices stay in bounds.
    {analysis -175}
    IF Value[ValueLength] = Terminator THEN
    {analysis +175}
        EXIT;
    END_IF;
END_FOR;

FOR SuffixLength := 0 TO UINT_TO_DINT(Param_Assertions.AssertionStringLength) DO
    // SA0175: Exact byte comparison; caller validates termination/capacity and indices stay in bounds.
    {analysis -175}
    IF Suffix[SuffixLength] = Terminator THEN
    {analysis +175}
        EXIT;
    END_IF;
END_FOR;

IF SuffixLength > ValueLength THEN
    RETURN;
END_IF;

SuffixStartIndex := ValueLength - SuffixLength;
FOR CharacterIndex := 0 TO SuffixLength - 1 DO
    // SA0175: Exact byte comparison; caller validates termination/capacity and indices stay in bounds.
    {analysis -175}
    IF Value[SuffixStartIndex + CharacterIndex] <> Suffix[CharacterIndex] THEN
    {analysis +175}
        RETURN;
    END_IF;
END_FOR;

TextEndsWith_String := TRUE;

END_FUNCTION

// ---- Framework/Assertions/POU/Utilities/TextStartsWith_String.TcPOU
{region 'Documentation'}
(*!
<summary>Exact prefix comparison without copies; an empty prefix matches. Caller supplies valid, stable references and content within the configured assertion capacity.</summary>
*)
{endregion}
FUNCTION INTERNAL TextStartsWith_String : BOOL //! TRUE when Value starts with Prefix; an empty Prefix matches.
VAR_IN_OUT CONSTANT
    Value : STRING(Param_Assertions.AssertionStringLength); //! Read-only source text; must be terminated within the configured capacity and stable during the call.
    Prefix : STRING(Param_Assertions.AssertionStringLength); //! Read-only prefix compared by code unit; an empty value matches in this helper.
END_VAR
VAR
    CharacterIndex : DINT;
END_VAR
VAR CONSTANT
    Terminator : BYTE := 0;
END_VAR

TextStartsWith_String := FALSE;

FOR CharacterIndex := 0 TO UINT_TO_DINT(Param_Assertions.AssertionStringLength) DO
    // SA0175: Exact byte comparison; caller validates termination/capacity and indices stay in bounds.
    {analysis -175}
    IF Prefix[CharacterIndex] = Terminator THEN
    {analysis +175}
        TextStartsWith_String := TRUE;
        RETURN;
    END_IF;

    // SA0175: Exact byte comparison; caller validates termination/capacity and indices stay in bounds.
    {analysis -175}
    IF Value[CharacterIndex] <> Prefix[CharacterIndex] THEN
    {analysis +175}
        RETURN;
    END_IF;
END_FOR;

END_FUNCTION

// ---- Framework/Assertions/POU/Utilities/TextEndsWith_WString.TcPOU
{region 'Documentation'}
(*!
<summary>Exact suffix comparison without copies; an empty suffix matches. Caller supplies valid, stable references and content within the configured assertion capacity.</summary>
*)
{endregion}
FUNCTION INTERNAL TextEndsWith_WString : BOOL //! TRUE when Value ends with Suffix; an empty Suffix matches.
VAR_IN_OUT CONSTANT
    Value : WSTRING(Param_Assertions.AssertionWStringLength); //! Read-only source text; must be terminated within the configured capacity and stable during the call.
    Suffix : WSTRING(Param_Assertions.AssertionWStringLength); //! Read-only suffix compared by code unit; an empty value matches in this helper.
END_VAR
VAR
    CharacterIndex : DINT;
    ValueLength : DINT;
    SuffixLength : DINT;
    SuffixStartIndex : DINT;
END_VAR
VAR CONSTANT
    Terminator : WORD := 0;
END_VAR

TextEndsWith_WString := FALSE;

FOR ValueLength := 0 TO UINT_TO_DINT(Param_Assertions.AssertionWStringLength) DO
    IF Value[ValueLength] = Terminator THEN
        EXIT;
    END_IF;
END_FOR;

FOR SuffixLength := 0 TO UINT_TO_DINT(Param_Assertions.AssertionWStringLength) DO
    IF Suffix[SuffixLength] = Terminator THEN
        EXIT;
    END_IF;
END_FOR;

IF SuffixLength > ValueLength THEN
    RETURN;
END_IF;

SuffixStartIndex := ValueLength - SuffixLength;
FOR CharacterIndex := 0 TO SuffixLength - 1 DO
    IF Value[SuffixStartIndex + CharacterIndex] <> Suffix[CharacterIndex] THEN
        RETURN;
    END_IF;
END_FOR;

TextEndsWith_WString := TRUE;

END_FUNCTION

// ---- Framework/Assertions/POU/Utilities/TextStartsWith_WString.TcPOU
{region 'Documentation'}
(*!
<summary>Exact prefix comparison without copies; an empty prefix matches. Caller supplies valid, stable references and content within the configured assertion capacity.</summary>
*)
{endregion}
FUNCTION INTERNAL TextStartsWith_WString : BOOL //! TRUE when Value starts with Prefix; an empty Prefix matches.
VAR_IN_OUT CONSTANT
    Value : WSTRING(Param_Assertions.AssertionWStringLength); //! Read-only source text; must be terminated within the configured capacity and stable during the call.
    Prefix : WSTRING(Param_Assertions.AssertionWStringLength); //! Read-only prefix compared by code unit; an empty value matches in this helper.
END_VAR
VAR
    CharacterIndex : DINT;
END_VAR
VAR CONSTANT
    Terminator : WORD := 0;
END_VAR

TextStartsWith_WString := FALSE;

FOR CharacterIndex := 0 TO UINT_TO_DINT(Param_Assertions.AssertionWStringLength) DO
    IF Prefix[CharacterIndex] = Terminator THEN
        TextStartsWith_WString := TRUE;
        RETURN;
    END_IF;

    IF Value[CharacterIndex] <> Prefix[CharacterIndex] THEN
        RETURN;
    END_IF;
END_FOR;

END_FUNCTION

// ---- Framework/EventBuffer/POU/EventBufferDiagConsumer.TcPOU
{region 'Documentation'}
(*!
<summary>Discards events for PLC-only lifecycle diagnosis; this is not an evaluated test run.</summary>
<description>
Call once per cycle after RunControl in the same task, including during initial Reset.
Supply the initialized buffer service and its actual one-based event storage. No other consumer
may acknowledge this epoch. The array is borrowed only for this call, never copied or retained.
Activation consumes immediately; subsequent batches follow ConsumeInterval without catch-up.
Disabled calls neither access the buffer nor clear held diagnostics. No events are evaluated.


HasError describes diagnostic consumption, not the test verdict. A batch attempt clears its previous batch/error state before work; a failing batch retains confirmed partial progress and reports Error. ResetDiagnostics clears observations only. Disabling resets the interval schedule, so the next valid activation consumes immediately; it does not reset the buffer or its epoch.
</description>
*)
{endregion}
FUNCTION_BLOCK EventBufferDiagConsumer
VAR_INPUT
    Enable : BOOL := FALSE; //! Enables event discarding; default FALSE. The first enabled call consumes immediately.
    Buffer : I_EventBuffer; //! Initialized service for the supplied Events array; no other consumer may acknowledge this epoch.
END_VAR
VAR_IN_OUT CONSTANT
    Events : ARRAY[*] OF ST_Event; //! Read-only physical ring storage belonging to Buffer; borrowed only for this call, not retained.
END_VAR
VAR
    FEnabled : BOOL;
    FMaxEventsPerCall : UINT := 32;
    FConsumeInterval : TIME := T#10ms;
    FIntervalTimer : Stopwatch;
    FDiscardedEventCount : ULINT;
    FLastBatchEventCount : UINT;
    FPeakPendingEventCount : UINT;
    FHasError : BOOL;
END_VAR
VAR_TEMP
    PendingStatus : ST_FifoStatus;
END_VAR

IF NOT Enable THEN
    FEnabled := FALSE;
    FIntervalTimer.Reset();
    RETURN;
END_IF;

IF Buffer = 0 THEN
    FHasError := TRUE;
    RETURN;
END_IF;

PendingStatus := Buffer.FifoStatus;
IF PendingStatus.ConfigError OR PendingStatus.IndexError
    OR (PendingStatus.BufferLength < 2)
    OR (PendingStatus.ElementCount >= PendingStatus.BufferLength) THEN
    FHasError := TRUE;
    RETURN;
END_IF;
FPeakPendingEventCount := MAX(FPeakPendingEventCount, PendingStatus.ElementCount);

IF FEnabled THEN
    FIntervalTimer.Update();
    IF NOT FIntervalTimer.IsValid THEN
        FHasError := TRUE;
        FIntervalTimer.Start();
        RETURN;
    END_IF;
    IF FIntervalTimer.ElapsedTime < FConsumeInterval THEN
        RETURN;
    END_IF;
END_IF;

FEnabled := TRUE;
ConsumeEvents(Events := Events);
FIntervalTimer.Start();

{region 'Documentation'}
(*!
<summary>Discards at most one bounded batch from the FIFO head; counts only confirmed deletions.</summary>
<description>
An invalid binding, range, sequence or rejected deletion stops this batch and sets HasError.
Buffer and Events must identify the same storage; equal dimensions alone cannot prove identity.
</description>
*)
{endregion}
METHOD PRIVATE ConsumeEvents
VAR_IN_OUT CONSTANT
    Events : ARRAY[*] OF ST_Event; //! Read-only one-based storage of Buffer, borrowed for this batch without copying or retention.
END_VAR
VAR
    FifoStatus : ST_FifoStatus;
    BufferStatus : ST_EventBufferStatus;
    BatchLimit : UINT;
    EntryNumber : UINT;
    HeadSequenceId : UDINT;
    DeleteSequenceId : UDINT;
END_VAR
VAR CONSTANT
    MaxDiscardedEventCount : ULINT := ULINT#18446744073709551615;
END_VAR
FLastBatchEventCount := 0;
FHasError := FALSE;
IF FMaxEventsPerCall = 0 THEN
    FHasError := TRUE;
    RETURN;
END_IF;

FifoStatus := Buffer.FifoStatus;
IF FifoStatus.ConfigError OR FifoStatus.IndexError
    OR (FifoStatus.BufferLength < 2)
    OR (LOWER_BOUND(Events, 1) <> 1)
    OR (UPPER_BOUND(Events, 1) <> UINT_TO_DINT(FifoStatus.BufferLength))
    OR (FifoStatus.ElementCount >= FifoStatus.BufferLength) THEN
    FHasError := TRUE;
    RETURN;
END_IF;

BatchLimit := MIN(FMaxEventsPerCall, FifoStatus.ElementCount);
FOR EntryNumber := 1 TO BatchLimit DO
    FifoStatus := Buffer.FifoStatus;
    IF FifoStatus.ConfigError OR FifoStatus.IndexError
        OR (FifoStatus.IndexOut < 1) OR (FifoStatus.IndexOut > FifoStatus.BufferLength) THEN
        FHasError := TRUE;
        RETURN;
    END_IF;
    IF FifoStatus.BufferEmpty THEN
        EXIT;
    END_IF;

    HeadSequenceId := Events[FifoStatus.IndexOut].SequenceId;
    BufferStatus := Buffer.Status;
    IF (HeadSequenceId = 0)
        OR (HeadSequenceId <= BufferStatus.DeletedSequenceId)
        OR (HeadSequenceId > BufferStatus.SequenceId) THEN
        FHasError := TRUE;
        RETURN;
    END_IF;

    DeleteSequenceId := HeadSequenceId;
    Buffer.ProcessDeleteRequest(SequenceId := DeleteSequenceId);
    BufferStatus := Buffer.Status;
    IF BufferStatus.DeletedSequenceId <> HeadSequenceId THEN
        FHasError := TRUE;
        RETURN;
    END_IF;

    FLastBatchEventCount := FLastBatchEventCount + 1;
    IF FDiscardedEventCount < MaxDiscardedEventCount THEN
        FDiscardedEventCount := FDiscardedEventCount + 1;
    END_IF;
END_FOR;
END_METHOD

{region 'Documentation'}
(*!
<summary>Minimum batch interval, default T#10ms. T#0ms consumes every call; no catch-up batches.</summary>
*)
{endregion}
{attribute 'monitoring' := 'call'}
PROPERTY PUBLIC ConsumeInterval : TIME //! Minimum batch interval, default T#10ms. T#0ms consumes every call; no catch-up batches.
GET // PUBLIC
ConsumeInterval := FConsumeInterval;
END_GET
SET // PUBLIC
FConsumeInterval := ConsumeInterval;
END_SET
END_PROPERTY

{region 'Documentation'}
(*!
<summary>Confirmed discarded events since ResetDiagnostics, saturating at ULINT maximum; independent of buffer epochs.</summary>
*)
{endregion}
{attribute 'monitoring' := 'call'}
PROPERTY PUBLIC DiscardedEventCount : ULINT //! Confirmed discarded events since ResetDiagnostics, saturating at ULINT maximum; independent of buffer epochs.
GET // PUBLIC
DiscardedEventCount := FDiscardedEventCount;
END_GET
END_PROPERTY

{region 'Documentation'}
(*!
<summary>Buffer observation, batch or time-base failure; retained until a batch succeeds or ResetDiagnostics is called.</summary>
*)
{endregion}
{attribute 'monitoring' := 'call'}
PROPERTY PUBLIC HasError : BOOL //! Buffer observation, batch or time-base failure; retained until a batch succeeds or ResetDiagnostics is called.
GET // PUBLIC
HasError := FHasError;
END_GET
END_PROPERTY

{region 'Documentation'}
(*!
<summary>Actual deletions in the last attempted batch, including partial failure; held between batches and while disabled.</summary>
*)
{endregion}
{attribute 'monitoring' := 'call'}
PROPERTY PUBLIC LastBatchEventCount : UINT //! Actual deletions in the last attempted batch, including partial failure; held between batches and while disabled.
GET // PUBLIC
LastBatchEventCount := FLastBatchEventCount;
END_GET
END_PROPERTY

{region 'Documentation'}
(*!
<summary>Maximum events per cyclic call, default 32. Zero is invalid and prevents consumption.</summary>
*)
{endregion}
{attribute 'monitoring' := 'call'}
PROPERTY PUBLIC MaxEventsPerCall : UINT //! Maximum events per cyclic call, default 32. Zero is invalid and prevents consumption.
GET // PUBLIC
MaxEventsPerCall := FMaxEventsPerCall;
END_GET
SET // PUBLIC
FMaxEventsPerCall := MaxEventsPerCall;
END_SET
END_PROPERTY

{region 'Documentation'}
(*!
<summary>Highest valid pre-consumption occupancy sampled on every enabled call since ResetDiagnostics; not only at batch intervals.</summary>
*)
{endregion}
{attribute 'monitoring' := 'call'}
PROPERTY PUBLIC PeakPendingEventCount : UINT //! Highest valid pre-consumption occupancy sampled on every enabled call since ResetDiagnostics; not only at batch intervals.
GET // PUBLIC
PeakPendingEventCount := FPeakPendingEventCount;
END_GET
END_PROPERTY

{region 'Documentation'}
(*!
<summary>Immediately clears only the three consumer statistics and error indication; no buffer or scheduling effects.</summary>
*)
{endregion}
METHOD PUBLIC ResetDiagnostics
FDiscardedEventCount := 0;
FLastBatchEventCount := 0;
FPeakPendingEventCount := 0;
FHasError := FALSE;
END_METHOD

END_FUNCTION_BLOCK

// ---- Framework/EventBuffer/POU/StateTransitionEvents/CreateTestCaseOrchestratorStateTransitionEvent.TcPOU
{region 'Documentation'}
(*!
<summary>Constructs a Test Case Orchestrator transition event without publishing it.</summary>
<description>
Name is the parent name; the appended .Orchestrator name uses the fixed event capacity.


This retained technical constructor is not called by the current owner-driven Orchestrator, which emits Framework error diagnostics rather than normal task/slot transitions. Its technical scope/name never supplies Full Owner completion evidence.
</description>
*)
{endregion}
FUNCTION CreateTestCaseOrchestratorStateTransitionEvent : ST_Event //! Constructed event value; not published. The publisher assigns SequenceId and Timestamp.
VAR_INPUT
    Name : STRING(GVL_Constants.NameLength); //! Parent's hierarchical name; the event name appends '.Orchestrator'.
    StateOld : E_State; //! Owner state before the reported or rejected transition.
    StateNew : E_State; //! Requested destination state recorded in the event; this function does not perform the transition.
END_VAR

CreateTestCaseOrchestratorStateTransitionEvent.SequenceId := 0;
CreateTestCaseOrchestratorStateTransitionEvent.Timestamp := 0;
CreateTestCaseOrchestratorStateTransitionEvent.OwnerScope := E_OwnerScope.TestCaseOrchestrator;
CreateTestCaseOrchestratorStateTransitionEvent.EventType := E_EventType.StateTransition;
CreateTestCaseOrchestratorStateTransitionEvent.Severity := E_EventSeverity.Info;
CreateTestCaseOrchestratorStateTransitionEvent.Name := CONCAT(STR1 := Name,
    STR2 := '.Orchestrator');
CreateTestCaseOrchestratorStateTransitionEvent.ResourceName := '';
CreateTestCaseOrchestratorStateTransitionEvent.State := StateNew;
CreateTestCaseOrchestratorStateTransitionEvent.Result := E_Result.NotEvaluated;
CreateTestCaseOrchestratorStateTransitionEvent.Message := CONCAT(STR1 := 'State transition ',
    STR2 := INT_TO_STRING(TO_INT(StateOld)));
CreateTestCaseOrchestratorStateTransitionEvent.Message := CONCAT(STR1 := CreateTestCaseOrchestratorStateTransitionEvent.Message,
    STR2 := ' -> ');
CreateTestCaseOrchestratorStateTransitionEvent.Message := CONCAT(STR1 := CreateTestCaseOrchestratorStateTransitionEvent.Message,
    STR2 := INT_TO_STRING(TO_INT(StateNew)));

END_FUNCTION

// ---- Framework/EventBuffer/POU/StateTransitionEvents/CreateTestSuiteOrchestratorStateTransitionEvent.TcPOU
{region 'Documentation'}
(*!
<summary>Constructs a Test Suite Orchestrator transition event without publishing it.</summary>
<description>
Name is the parent name; the appended .Orchestrator name uses the fixed event capacity.


This retained technical constructor is not called by the current owner-driven Orchestrator, which emits Framework error diagnostics rather than normal task/slot transitions. Its technical scope/name never supplies Full Owner completion evidence.
</description>
*)
{endregion}
FUNCTION CreateTestSuiteOrchestratorStateTransitionEvent : ST_Event //! Constructed event value; not published. The publisher assigns SequenceId and Timestamp.
VAR_INPUT
    Name : STRING(GVL_Constants.NameLength); //! Parent's hierarchical name; the event name appends '.Orchestrator'.
    StateOld : E_State; //! Owner state before the reported or rejected transition.
    StateNew : E_State; //! Requested destination state recorded in the event; this function does not perform the transition.
END_VAR

CreateTestSuiteOrchestratorStateTransitionEvent.SequenceId := 0;
CreateTestSuiteOrchestratorStateTransitionEvent.Timestamp := 0;
CreateTestSuiteOrchestratorStateTransitionEvent.OwnerScope := E_OwnerScope.TestSuiteOrchestrator;
CreateTestSuiteOrchestratorStateTransitionEvent.EventType := E_EventType.StateTransition;
CreateTestSuiteOrchestratorStateTransitionEvent.Severity := E_EventSeverity.Info;
CreateTestSuiteOrchestratorStateTransitionEvent.Name := CONCAT(STR1 := Name,
    STR2 := '.Orchestrator');
CreateTestSuiteOrchestratorStateTransitionEvent.ResourceName := '';
CreateTestSuiteOrchestratorStateTransitionEvent.State := StateNew;
CreateTestSuiteOrchestratorStateTransitionEvent.Result := E_Result.NotEvaluated;
CreateTestSuiteOrchestratorStateTransitionEvent.Message := CONCAT(STR1 := 'State transition ',
    STR2 := INT_TO_STRING(TO_INT(StateOld)));
CreateTestSuiteOrchestratorStateTransitionEvent.Message := CONCAT(STR1 := CreateTestSuiteOrchestratorStateTransitionEvent.Message,
    STR2 := ' -> ');
CreateTestSuiteOrchestratorStateTransitionEvent.Message := CONCAT(STR1 := CreateTestSuiteOrchestratorStateTransitionEvent.Message,
    STR2 := INT_TO_STRING(TO_INT(StateNew)));

END_FUNCTION
